(* IEC 61131-3 sources: daoli-st-library/DL_Base (part 7) *)

(* ---- FC_DL_RorEx.st ---- *)
(*==============================================================================
 * 组件名称 (Component)  : FC_DL_RorEx
 * 所属子库 (Sublibrary) : DL_Base
 * 当前版本 (Version)    : 1.0.0
 * 兼容性   (Platform)   : CODESYS 3.5 / TwinCAT 3 / 汇川 InoProShop / Machine Expert
 *                         仅依赖 Standard.library 的 SHL / SHR 内建函数，
 *                         循环语义由移位合成显式构造，无厂商 ROR 方言依赖
 * 功能一句话 (Summary)  : 循环右移防御包装：移位量对位宽取模归一后再循环，
 *                         杜绝平台相关行为，循环位不丢。
 * 功能描述 (Function)   : 对被移位位串按移位量 nN 循环右移。归一策略写死：
 *                         nN 先 MOD 32 归一到 0 到 31（nN 为 USINT 天然非负，
 *                         禁用 MOD 对负数的平台歧义取余的前提由类型系统保证）；
 *                         归一后 nN = 0 直接返回原值（整圈等价于不动，不置码）；
 *                         归一后 1 到 31 用「右移 nN OR 左移 (32 − nN)」位合成
 *                         构造循环语义，两个合成移位量均严格落在 1 到 31 安全域。
 * 溯源     (Origin)     : IEC 61131-3 标准语义的道莅防御性实现
 *                         （接口语义由 IEC 61131-3 定义，clean-room 重写，
 *                         参考公开标准条款）
 * 支持位宽 (Width Note) : 本件按 DWORD（32 位）主类型实现，仅支持 32 位位串；
 *                         BYTE / WORD 调用方先显式转换到 DWORD 后调用，再按需
 *                         截回原位宽（头注释显式声明，不做 ANY_BIT 泛型）。
 * 类型裁定 (Type Note)  : 码位段 16#0001_xxxx 为全库共享 32 位段，WORD 容量不足，
 *                         故 uDiag 采用 UDINT 承载（与库内 uErrorId : UDINT 惯例一致）
 * 依赖     (Depends)    : 无 DL_ 内部依赖；Standard.library: SHL / SHR
 * 红线自检 (Redline)    : R1 ✓ 零全局变量与外部变量引用 ｜ R2 ✓ 零物理 IO 地址直写
 *                         R3 ✓ 纯 IEC 61131-3 ｜ R4 ✓ 移位量 MOD 归一（合成移位
 *                         量恒在 1 到 31 安全域）｜ R5 ✓ 全变量中英双语同行注释
 *                         R6 N/A（纯函数，无 CASE/ENUM 状态机，按批 1 口径标 N/A）
 *                         R7 N/A（FC 为纯函数，无实例调用，头注释显式说明）
 * 防御行为声明 (Defense): ① 归一先行：nN ≥ 32 时先 MOD 32 归一并置信息码
 *                           16#0001_0159（已归一提示），归一后绝不出现 ≥ 位宽
 *                           的移位量，杜绝平台对超宽循环移位的歧义行为；
 *                         ② nN 为 USINT 类型天然非负，MOD 只作用于非负域，
 *                           负数取余的平台歧义（如商向零取整方向不一）从类型
 *                           系统层面被排除，该前提已在头注释写死；
 *                         ③ 归一后 nN = 0 直接返回原值且不置码（整圈无事件）；
 *                         ④ 位合成用「SHR(uIn, nN) OR SHL(uIn, 32 − nN)」，
 *                           nN 归一后为 1 到 31，故 32 − nN 恒为 1 到 31，
 *                           两个移位量均不触碰「移位量 = 位宽」禁区，循环位不丢；
 *                         ⑤ 32（位宽）提为只读常量，禁魔法数。
 * 修订历史 (Revision)   :
 *   2026-11-16  v1.0.0  首版入库（R14 批 3 · T0 快车道）
 *============================================================================*)
FUNCTION FC_DL_RorEx : DWORD
VAR_INPUT
    uIn : DWORD;   // 被循环移位位串 [位] / Bit string to be rotated
    nN  : USINT;   // 移位量 [bit]，USINT 天然非负，MOD 仅作用于非负域 / Shift amount [bit], USINT is non-negative, MOD applied on the non-negative domain only
END_VAR
VAR_OUTPUT
    uDiag : UDINT; // 诊断字，16#0001_0159=移位量已 MOD 32 归一，0=无事件 / Diag word, 16#0001_0159=shift amount reduced by MOD 32, 0=no event
END_VAR
VAR
    nNorm : USINT; // 归一后移位量 [bit]，域 0 到 31 / Normalized shift amount [bit], range 0 to 31
END_VAR
VAR CONSTANT
    DL_RR_WIDTH : USINT := 32;  // 位宽常量 [bit]，MOD 归一与合成移位共用 / Width constant [bit], shared by MOD normalization and composite shifts
END_VAR

(*------------------------------------------------------------------------------
 * 段 1｜输出与诊断预置：先归零，任何路径都不会留下脏诊断
 *      Pre-set the output and diag so no path ever leaves a stale diag
 *-----------------------------------------------------------------------------*)
FC_DL_RorEx := 16#0000_0000;   // 返回值预置全零 [位串] / Preset return value to all zero
uDiag       := 16#0000_0000;   // 诊断字预置无事件 / Preset diag word to no event
nNorm       := 0;              // 归一移位量预置 [bit] / Preset normalized shift to zero [bit]

(*------------------------------------------------------------------------------
 * 段 2｜移位量归一（防御声明①②）：nN MOD 32 归一到 0 到 31；
 *      nN 为 USINT 非负域，MOD 结果即数学取模，无负数取余歧义；
 *      nN ≥ 32 置信息码提示已归一（归一是正常防御行为，非故障）
 *      Shift-amount normalization (defense notes 1 and 2): nN MOD 32 reduces
 *      to 0 to 31; a reduction raises the informational code, not a fault
 *-----------------------------------------------------------------------------*)
IF nN >= DL_RR_WIDTH THEN
    nNorm := nN MOD DL_RR_WIDTH;   // 超宽归一：MOD 32 取模 [bit] / Oversized normalization: MOD 32 [bit]
    uDiag := 16#0001_0159;         // 信息码：移位量已 MOD 32 归一 / Informational: shift amount reduced by MOD 32
ELSE
    nNorm := nN;                   // 域内直通 [bit] / In-domain pass-through [bit]
END_IF

(*------------------------------------------------------------------------------
 * 段 3｜循环移位主体（防御声明③④）：归一后 0 整圈直通原值；
 *      1 到 31 用右移与左移位合成，合成移位量恒在安全域，循环位不丢
 *      Rotation body (defense notes 3 and 4): normalized zero returns as is;
 *      one to thirty one composes SHR and SHL, both amounts stay in the safe
 *      domain so no bit is ever lost
 *-----------------------------------------------------------------------------*)
IF nNorm = 0 THEN
    FC_DL_RorEx := uIn;   // 整圈（或 0 位）等价于原值直通 [位串] / A full turn (or zero shift) returns the input unchanged
ELSE
    FC_DL_RorEx := SHR(uIn, nNorm) OR SHL(uIn, DL_RR_WIDTH - nNorm);   // 位合成循环右移 [位串] / Composite rotate right
END_IF
END_FUNCTION

(* ---- FC_DL_RorLwordEx.st ---- *)
(*
    FC_DL_RorLwordEx —— LWORD 循环右移（MOD 64 归一）
    ------------------------------------------------------------------
    分类      : DL_Base / BitString
    前缀      : FC_DL_
    版本      : 1.0.0
    溯源      : IEC 61131-3 标准语义的道莅防御性实现
                （接口语义由 IEC 61131-3 定义，内部委托平台内建 ROR，
                  外围统一错误码 / 钳位 / 双语文档；clean-room 重写，
                  未复制任何闭源厂商源码，参考实现仅限 MIT/Apache 许可）
    平台      : 纯 IEC 61131-3，CODESYS / TwinCAT / InoProShop 通用
    作者      : 道莅代码库 · PLC编程专家（R17）
    ------------------------------------------------------------------
    功能说明  : LWORD 位串循环右移防御包装：移位量 nN 大于等于 64（位宽）时按 MOD 64 归一，
                并置信息级 16#0001_020C（与循环左移件同口径，与左移/右移件的「超宽置零」刻意相反）；
                归一后移位量为 0 时直接输出原值，不调用内建 ROR；
                域内委托平台内建 ROR，不重实现移位内核；
                MOD 除子为常量 64（编译期恒非零），结构性满足除法前判除子非零红线；
                钳位方向：移位量按位宽取模归一（0~63），结果位宽严格保持 64 位。
    错误码    : 16#0001_020C 移位量 ≥ 64（位宽），已按 MOD 64 归一——信息级，正常防御
                16#0001_020D 预留禁用（信息级，不得挪用）
                16#0001_0300 预留禁用（故障级，不得挪用）
                16#0001_0301 预留禁用（故障级，不得挪用）
                16#0001_0302 预留禁用（故障级，不得挪用）
    状态机    : R6 标注 N/A —— 本组件为纯函数无顺序状态机，无 CASE 可写，非法状态不可能出现，故以本节说明替代 ELSE 兜底
    修订记录  : 2026-11-16 v1.0.0 首次入库（R17）
*)
FUNCTION FC_DL_RorLwordEx : LWORD
VAR_INPUT
    uIn : LWORD; // 被循环移位位串 [位] / bit string to be rotated [bit]
    nN  : USINT; // 循环移位量 [bit]，USINT 天然非负，范围 0~255 / rotate amount [bit], USINT is non-negative by type, range 0..255
END_VAR
VAR_OUTPUT
    eErr   : UDINT; // 错误码，0=正常 / error id, 0=ok
    bError : BOOL;  // 是否出错，eErr 非 0 时为 TRUE / error flag, TRUE when eErr is nonzero
    bValid : BOOL;  // 输出是否有效可用 / output valid flag
END_VAR
VAR CONSTANT
    DL_LW_WIDTH : USINT := 64; // LWORD 位宽常量，兼作 MOD 除子（编译期恒非零） [bit] / LWORD width constant, also the MOD divisor, never zero [bit]
END_VAR
VAR
    nShift : USINT; // 归一后的实际移位量 0~63 [bit] / normalized shift amount 0..63 [bit]
END_VAR

// 段 1｜输出与错误状态预置 / segment 1, preset output and error status
FC_DL_RorLwordEx := uIn; // 输出预置为原值（零移位等价语义），任何路径不留脏值 [位串] / preset output to the input, the zero-shift identity, no stale value on any path [bit string]
eErr   := 0;     // 预置无错误 / preset no error
bError := FALSE; // 预置无故障（本件无故障级路径） / preset no fault, no fault-level path here
bValid := FALSE; // 预置输出无效，通过归一后置位 / preset invalid, set TRUE after normalization

// 段 2｜移位量归一（MOD 位宽） / segment 2, shift amount normalization (modulo width)
nShift := nN; // 默认按原移位量直通 [bit] / pass the original shift amount through by default [bit]
IF nN >= DL_LW_WIDTH THEN // 循环移位对位宽取模仍等价，故归一而非置零 [bit] / rotate modulo the width stays equivalent, so normalize instead of zeroing [bit]
    nShift := nN MOD DL_LW_WIDTH; // 除子为编译期常量 64，恒非零 [bit] / divisor is the compile-time constant 64, never zero [bit]
    eErr := 16#0001_020C;         // 信息级：移位量已归一，正常防御 / info level: shift amount normalized, normal defence
ELSE
    eErr := 0;                    // 未超宽，无记录 / not oversized, nothing recorded
END_IF

// 段 3｜零移位量与域内委托循环移位（末段） / segment 3, zero-shift pass-through and in-domain delegated rotate (final)
IF nShift = 0 THEN
    FC_DL_RorLwordEx := uIn; // 零移位量直接输出原值，规避内建 ROR 的平台差异 [位串] / zero shift passes the input through, avoiding platform differences of built-in ROR [bit string]
ELSE
    FC_DL_RorLwordEx := ROR(uIn, nShift); // 域内委托平台内建 ROR，不重实现移位内核 [位串] / in-domain delegate to built-in ROR, shift kernel not re-implemented [bit string]
END_IF
bError := FALSE; // 信息级不置故障 / info level never raises fault
bValid := TRUE;  // 归一后输出有效可用 / output is valid after normalization
END_FUNCTION

(* ---- FC_DL_SaturateDiv.st ---- *)
(*
  ==================================================================
  组件名 Component  : FC_DL_SaturateDiv
  分类   Category   : DL_Base
  前缀   Naming     : FC_DL_ ｜ b/n/u/f/t/e/st 类型前缀制（R265）
  码位   Code ID    : 16#0001_0647（信息级）｜ 16#0001_0648 / 0649 / 064A（故障级）
  版本   Version    : 1.0.0
  复杂度 Complexity  : 中
  功能   Purpose    : LINT 宽域饱和除法：nOut = clamp(nNum ÷ nDen, nLo, nHi)，判据有序
                      （除零 → MIN÷-1 → 正常除 → 域钳），整数商向零截断。
  开源溯源 Origin    : IEC 61131-3 标准语义的道莅防御性实现（clean-room，无第三方代码行）
  许可证 License    : MIT
  参考   Reference  : IEC 61131-3:2013 §6.6.2 算术运算符（整数除法，商向零截断）
  平台   Platform   : 纯 IEC 61131-3（仅四则与比较），CODESYS / TwinCAT 3 / InoProShop 通用
  依赖   Depends    : 仅 Standard.library（无库调用）
  分工声明 Split     : FC_DL_DivDintSafeChk 为「安全除 + 商出口 + 布尔返回」的判据件
                      （DINT 域、无钳位域）；FC_DL_DivLrealSafe 为浮点域安全除；
                      本件为宽域（LINT）饱和除，带钳位域与三段标志。三者边界：
                      需要「除零仅判不钳」用前者，需要「浮点除法」用中者，
                      需要「整数宽域 + 钳位域 + 溢出标志」用本件（R216 双向互引）。
  归属 Ownership     : 本件无 TYPE 声明，全部引脚为 IEC 标准原生类型。
  ------------------------------------------------------------------
  边界 Boundary     :
                      一 判据严格有序：① 除数为零 → 早退（禁走钳位，钳位会把非法
                         结果伪装成合法边界）；② MIN ÷ -1 → 溢出钳 nHi；③ 正常除；
                         ④ 结果钳域 [nLo, nHi]；
                      二 商向零截断（IEC 语义）：-7 ÷ 2 = -3 而非 -4；本件不做四舍五入，
                         工程舍入口径归 FC_DL_RoundSat，有效位舍入归 FC_DL_RoundSigFigs；
                      三 nLo > nHi 判组态故障并返回 FALSE（与 FC_DL_SaturateMul、
                         FC_DL_RealToIntSat 同口径，三件一致，禁静默交换）；
                      四 纯函数：无记忆量、无定时器、无边沿实例，每调用重算。
  错误码 Codes      :
    16#0001_0647【信息级】结果被域 [nLo, nHi] 钳位（未溢出、未除零，bValid = TRUE）
    16#0001_0648【故障级】除数为零（nOut = 0，bValid = FALSE，早退不走钳位）
    16#0001_0649【故障级】MIN ÷ -1 溢出（nOut 钳 nHi，bOvF = TRUE）
    16#0001_064A【故障级】组态非法 nLo > nHi（判故障返回 FALSE，nOut = 0）
  码位反证 Note     :
    0648 不可并入 0647：除零结果与钳位结果在数值出口上同为边界值或零，上游无法由
    nOut 与 bClamped 组合区分「输入非法」与「输入合法但被限幅」，两码必需（R90）。
  验收 Acceptance   :
    算法已证（脚本）：未跑 ｜ 编译器已证（三平台）：未跑
    V1 5 ÷ 0 → 0、bDivZero = TRUE、bValid = FALSE、码 0648（不走钳位）
    V2 MIN ÷ -1 → nHi、bOvF = TRUE、码 0649
    V3 MIN ÷ 1 → MIN 精确
    V4 1 ÷ MIN → 0，bClamped = FALSE（未触钳位，仅截断）
    V5 -7 ÷ 2 → -3（向零截断，非 -4）
    V6 nLo > nHi → 码 064A、返回 FALSE
    V7 100 ÷ 3 = 33（截断）、域 [0, 20] → bClamped = TRUE、码 0647、bValid = TRUE
    V8 MIN ÷ -3 → 正常除（除子非 -1）不溢出
  修订记录 Revision  :
    2026-11-21  v1.0.0  R62 首版（批 1 · 序号 2）
  ==================================================================
*)
FUNCTION FC_DL_SaturateDiv : BOOL
VAR_INPUT
    nNum : LINT; // 被除数 [−]，完整 LINT 域 / the dividend over the full LINT domain
    nDen : LINT; // 除数 [−]，零为非法（判故障）/ the divisor, zero is illegal and raises a fault
    nLo  : LINT; // 输出钳位域下界 [−] / the output clamp lower bound
    nHi  : LINT; // 输出钳位域上界 [−] / the output clamp upper bound
END_VAR
VAR_OUTPUT
    nOut     : LINT;  // 钳位后商 [−] / the clamped quotient
    bDivZero : BOOL;  // 除数为零 [-] / the divisor is zero
    bOvF     : BOOL;  // 溢出发生（MIN ÷ -1）[-] / an overflow happened on MIN divided by minus one
    bClamped : BOOL;  // 钳位生效（含纯域钳）[-] / the clamp took effect, domain clamp included
    bValid   : BOOL;  // 输出可用（除零与组态故障为 FALSE）[-] / the output is usable
    eErr     : UDINT; // 错误码，0 = 正常 / the error code, zero is ok
    bError   : BOOL;  // 故障标志，故障级码同拍置位（R45 配对）/ the fault flag, raised with a fault level code
END_VAR
VAR
    liQuot : LINT := 0; // 域内商中间量 [−] / the in-domain quotient intermediate
END_VAR  // R64 结构补齐：VAR 段缺失的 END_VAR（门禁机械修复）
VAR CONSTANT
    DL_SDIV_MAX : LINT := 9223372036854775807;      // LINT 可表达上界 [−]，独立命名不与乘法件冲突 / the expressible LINT ceiling under its own name
    DL_SDIV_MIN : LINT := -9223372036854775807 - 1; // LINT 可表达下界 [−]，以上界相反数减一表达 / the expressible LINT floor written as the negated ceiling minus one
    DL_SDIV_ZERO : LINT := 0;                       // 有符号零常量 [−] / the signed zero constant
    DL_SDIV_NEG1 : LINT := -1;                      // 负一常量 [−]，MIN ÷ -1 判据用 / the minus one constant for the MIN divided by minus one criterion
END_VAR

// 段 1｜返回值与全部出口预置安全值（R45 四段式第一段）/ segment 1, preset every outlet to its safe value
FC_DL_SaturateDiv := FALSE; // 返回值预置假 / preset the return false
nOut := DL_SDIV_ZERO; // 结果预置零 [−] / preset the quotient zero
bDivZero := FALSE; // 除零标志预置假 / preset the divide by zero flag false
bOvF := FALSE; // 溢出标志预置假 / preset the overflow flag false
bClamped := FALSE; // 钳位标志预置假 / preset the clamp flag false
bValid := FALSE; // 可用标志预置假，过闸后置位 / preset the validity false, raised after the gates
eErr := 16#0000_0000; // 错误码预置正常 / preset the code to ok
bError := FALSE; // 故障标志预置假 / preset the fault flag false
liQuot := DL_SDIV_ZERO; // 商中间量清零 [−] / clear the quotient intermediate

// 段 2｜组态域闸：nLo > nHi 判故障早退（边界三，三件同口径）/ segment 2, the configuration gate, a reversed domain is a fault
IF nLo > nHi THEN // 钳位域反序 / the clamp domain is reversed
    eErr := 16#0001_064A; // 故障级：组态非法 nLo > nHi / fault grade, the reversed clamp domain
    bError := TRUE; // 同拍置故障标志（R45 配对）/ raise the fault flag on the same scan
    bValid := FALSE; // 输出不可用 / the output is not usable
    nOut := DL_SDIV_ZERO; // 确定缺省值零 [−] / the deterministic default of zero
    RETURN; // 早退 / early return
END_IF

// 段 3｜判据①除数为零：早退，绝不行钳位（边界一，钳位会把非法伪装成合法边界）/ segment 3, the divisor zero gate, clamped never runs
IF nDen = DL_SDIV_ZERO THEN // 除数为零 / the divisor is zero
    bDivZero := TRUE; // 置除零标志 / raise the divide by zero flag
    nOut := DL_SDIV_ZERO; // 确定缺省值零 [−] / the deterministic default of zero
    eErr := 16#0001_0648; // 故障级：除数为零 / fault grade, the divisor is zero
    bError := TRUE; // 同拍置故障标志（R45 配对）/ raise the fault flag on the same scan
    bValid := FALSE; // 输出不可用 / the output is not usable
    RETURN; // 早退，不做任何除法与钳位 / early return without any division or clamping
END_IF

// 段 4｜判据②MIN ÷ -1 溢出（MIN 的绝对值不可表示，先除必回绕）/ segment 4, the MIN divided by minus one overflow
IF (nNum = DL_SDIV_MIN) AND (nDen = DL_SDIV_NEG1) THEN // 极限组合 / the limit combination
    bOvF := TRUE; // 置溢出标志（禁回绕成 MIN）/ raise the overflow flag instead of wrapping to MIN
    bClamped := TRUE; // 钳位已生效 / the clamp took effect
    nOut := nHi; // 正溢出按符号钳上界 [−] / a positive overflow clamps to the upper bound by sign
    eErr := 16#0001_0649; // 故障级：MIN ÷ -1 溢出 / fault grade, the MIN divided by minus one overflow
    bError := TRUE; // 同拍置故障标志（R45 配对）/ raise the fault flag on the same scan
    bValid := FALSE; // 输出不可用 / the output is not usable
    RETURN; // 早退 / early return
END_IF

// 段 5｜判据③正常除：整数商向零截断（边界二，IEC 语义，-7 ÷ 2 = -3）/ segment 5, the normal division with the quotient truncated toward zero
IF nNum = DL_SDIV_ZERO THEN // 零被除数：商确为零，免一次除法 / a zero dividend gives an exact zero quotient, no division needed
    liQuot := DL_SDIV_ZERO; // 商为零 [−] / the quotient is zero
ELSE // 非零被除数才真除（除子已在段 3 证非零）/ the real division only for a nonzero dividend, the divisor is proven nonzero
    liQuot := nNum / nDen; // 向零截断（-7 ÷ 2 = -3，非 -4）[−] / truncated toward zero, minus seven over two gives minus three
END_IF

// 段 6｜判据④统一域钳（零被除数与正常除共用同一出口，R94）/ segment 6, the unified domain clamp shared by both paths
IF liQuot > nHi THEN // 超上界 / above the ceiling
    nOut := nHi; // 钳上界 [−] / clamp to the ceiling
    bClamped := TRUE; // 置钳位标志 / raise the clamp flag
ELSIF liQuot < nLo THEN // 超下界 / below the floor
    nOut := nLo; // 钳下界 [−] / clamp to the floor
    bClamped := TRUE; // 置钳位标志 / raise the clamp flag
ELSE // 域内 / inside the domain
    nOut := liQuot; // 直出商 [−] / pass the quotient through
END_IF

// 段 7｜信息级钳位码与可用位（纯域钳不置 bError，R285）/ segment 7, the informational clamp code without a fault flag
IF bClamped THEN // 发生纯域钳 / a pure domain clamp happened
    eErr := 16#0001_0647; // 信息级：结果被域钳位 / informational, the result was clamped to the domain
END_IF
bValid := TRUE; // 域内或钳位输出均可用 / an in-domain or clamped output is usable
FC_DL_SaturateDiv := TRUE; // 返回成功 / return success
END_FUNCTION

(* ---- FC_DL_SaturateMul.st ---- *)
(*
  ==================================================================
  组件名 Component  : FC_DL_SaturateMul
  分类   Category   : DL_Base
  前缀   Naming     : FC_DL_ ｜ b/n/u/f/t/e/st 类型前缀制（R265）
  码位   Code ID    : 16#0001_0644（信息级）｜ 16#0001_0645（故障级）｜ 16#0001_0646（故障级）
  版本   Version    : 1.0.0
  复杂度 Complexity  : 中
  功能   Purpose    : LINT 宽域饱和乘法：nOut = clamp(nA × nB, nLo, nHi)，溢出前判定，
                      bOvF（溢出）与 bClamped（钳位已生效）两标志语义可分。
  开源溯源 Origin    : IEC 61131-3 标准语义的道莅防御性实现（clean-room，无第三方代码行）
  许可证 License    : MIT
  参考   Reference  : IEC 61131-3:2013 §6.6.2 算术运算符（整数乘法）与 §6.6.5 类型转换语义
  平台   Platform   : 纯 IEC 61131-3（仅四则与比较），CODESYS / TwinCAT 3 / InoProShop 通用
  依赖   Depends    : 仅 Standard.library（无库调用）
  分工声明 Split     : 与 FC_DL_SaturateAdd（加）/ FC_DL_SaturateSub（减）构成「加/减/乘」
                      三件族，除法则由 FC_DL_SaturateDiv 承载；FC_DL_SaturateAdd 未覆盖
                      乘法（其模式枚举只有加与减），故本件不可省（R216 双向互引）。
  归属 Ownership     : 本件无 TYPE 声明，全部引脚为 IEC 标准原生类型。
  ------------------------------------------------------------------
  边界 Boundary     :
                      一 溢出前判定（禁先乘后判）：按四个象限分别与「域上界 ÷ 另一因子」
                         比较，比较式内只出现除法，不出现裸乘法，浮点无关、全整数精确；
                      二 MIN × -1 单独直判：MIN 的绝对值不可表示，先乘必回绕成 MIN 而
                         令「结果 < 0」误判为负溢出，故本组合在乘法之前直接判正溢出；
                      三 零因子优先：nA = 0 或 nB = 0 时积恒为 0，不做任何除法预判
                         （同时消灭预判式里的除零路径）；
                      四 nLo > nHi 判组态故障并返回 FALSE（与 FC_DL_SaturateDiv、
                         FC_DL_RealToIntSat 同口径，三件一致，禁静默交换）；
                      五 溢出与域钳两标志可分：溢出 → bOvF = TRUE 且 nOut 直达 nHi/nLo；
                         未溢出仅域钳 → bClamped = TRUE 且 bOvF = FALSE；
                      六 纯函数：无记忆量、无定时器、无边沿实例，每调用重算。
  错误码 Codes      :
    16#0001_0644【信息级】结果被域 [nLo, nHi] 钳位（未溢出，bClamped = TRUE，bValid = TRUE）
    16#0001_0645【故障级】乘法溢出（bOvF = TRUE，nOut 已按积符号钳到 nHi 或 nLo）
    16#0001_0646【故障级】组态非法 nLo > nHi（判故障返回 FALSE，nOut = 0）
  码位反证 Note     :
    0644 与 0645 不可合并：溢出与域钳在「结果数值」上不可观测区分（两者都输出边界值），
    仅靠返回值加 bValid 也无法分解（两者 bValid 不同，但 bOvF 语义才是上游限幅判据），
    故两码必需（R90 反证句：现有输出组合无法唯一还原该场景）。
  验收 Acceptance   :
    算法已证（脚本）：未跑 ｜ 编译器已证（三平台）：未跑
    V1 MAX × 2 → nOut = nHi、bOvF = TRUE、码 0645
    V2 MIN × -1 → nOut = nHi、bOvF = TRUE（禁回绕成 MIN）
    V3 MIN × 0 → 0 且 bOvF = FALSE
    V4 MIN × 1 → MIN 精确（无溢出、无钳位）
    V5 -3 × 5 → -15 精确
    V6 nLo > nHi → 码 0646、bError = TRUE、返回 FALSE
    V7 nLo = nHi = 100、积 = 200 → bClamped = TRUE 且 bOvF = FALSE（两标志可分）
    V8 nA = 0、nB = MIN → 0（零因子早于预判，无除零）
  修订记录 Revision  :
    2026-11-21  v1.0.0  R62 首版（批 1 · 序号 1）
  ==================================================================
*)
FUNCTION FC_DL_SaturateMul : BOOL
VAR_INPUT
    nA   : LINT; // 被乘数 [−]，完整 LINT 域 / the multiplicand over the full LINT domain
    nB   : LINT; // 乘数 [−]，完整 LINT 域 / the multiplier over the full LINT domain
    nLo  : LINT; // 输出钳位域下界 [−] / the output clamp lower bound
    nHi  : LINT; // 输出钳位域上界 [−] / the output clamp upper bound
END_VAR
VAR_OUTPUT
    nOut     : LINT;  // 钳位后结果 [−] / the clamped product
    bOvF     : BOOL;  // 乘法溢出发生（钳位已生效）[-] / a multiplicative overflow happened
    bClamped : BOOL;  // 钳位生效（含纯域钳，未溢出）[-] / the clamp took effect, domain clamp included
    bValid   : BOOL;  // 输出可用（溢出与组态故障为 FALSE）[-] / the output is usable
    eErr     : UDINT; // 错误码，0 = 正常 / the error code, zero is ok
    bError   : BOOL;  // 故障标志，故障级码同拍置位（R45 配对）/ the fault flag, raised with a fault level code
END_VAR
VAR
    liProd : LINT := 0; // 域内乘积中间量 [−] / the in-domain product intermediate
END_VAR  // R64 结构补齐：VAR 段缺失的 END_VAR（门禁机械修复）
VAR CONSTANT
    DL_SMUL_MAX : LINT := 9223372036854775807;      // LINT 可表达上界 [−]，即 2^63−1 / the expressible LINT ceiling, two to the sixty third minus one
    DL_SMUL_MIN : LINT := -9223372036854775807 - 1; // LINT 可表达下界 [−]，以上界相反数减一表达，防字面量解析溢出 / the expressible LINT floor, written as the negated ceiling minus one to avoid a literal parse overflow
    DL_SMUL_ZERO : LINT := 0;                       // 有符号零常量 [−]，避免裸字面量 / the signed zero constant
    DL_SMUL_NEG1 : LINT := -1;                      // 负一常量 [−]，MIN × -1 判据用 / the minus one constant for the MIN times minus one criterion
END_VAR

// 段 1｜返回值与全部出口预置安全值（R45 四段式第一段）/ segment 1, preset every outlet to its safe value
FC_DL_SaturateMul := FALSE; // 返回值预置假 / preset the return false
nOut := DL_SMUL_ZERO; // 结果预置零 [−] / preset the product zero
bOvF := FALSE; // 溢出标志预置假 / preset the overflow flag false
bClamped := FALSE; // 钳位标志预置假 / preset the clamp flag false
bValid := FALSE; // 可用标志预置假，过闸后置位 / preset the validity false, raised after the gates
eErr := 16#0000_0000; // 错误码预置正常 / preset the code to ok
bError := FALSE; // 故障标志预置假 / preset the fault flag false
liProd := DL_SMUL_ZERO; // 乘积中间量清零 [−] / clear the product intermediate

// 段 2｜组态域闸：nLo > nHi 判故障早退（边界四，三件同口径）/ segment 2, the configuration gate, a reversed domain is a fault
IF nLo > nHi THEN // 钳位域反序 / the clamp domain is reversed
    eErr := 16#0001_0646; // 故障级：组态非法 nLo > nHi / fault grade, the reversed clamp domain
    bError := TRUE; // 同拍置故障标志（R45 配对）/ raise the fault flag on the same scan
    bValid := FALSE; // 输出不可用 / the output is not usable
    nOut := DL_SMUL_ZERO; // 确定缺省值零 [−] / the deterministic default of zero
    RETURN; // 早退，不再触碰乘法 / early return, the multiplication is never touched
END_IF

// 段 3｜零因子优先：积恒为零，且消灭后续预判式的除零路径（边界三）/ segment 3, the zero factor comes first and removes every division by zero
IF (nA = DL_SMUL_ZERO) OR (nB = DL_SMUL_ZERO) THEN // 任一因子为零 / either factor is zero
    liProd := DL_SMUL_ZERO; // 积确定为零 [−] / the product is exactly zero
ELSE // 双因子非零才做溢出预判 / the overflow pre-check runs only with two nonzero factors
    // 段 4｜MIN × -1 直判正溢出（边界二）：MIN 绝对值不可表示，先乘会回绕成 MIN / segment 4, the direct check of MIN times minus one
    IF ((nA = DL_SMUL_MIN) AND (nB = DL_SMUL_NEG1)) OR ((nB = DL_SMUL_MIN) AND (nA = DL_SMUL_NEG1)) THEN // 极限组合 / the limit combination
        bOvF := TRUE; // 置溢出标志（禁回绕成 MIN）/ raise the overflow flag instead of wrapping to MIN
        bClamped := TRUE; // 钳位已生效 / the clamp took effect
        nOut := nHi; // 正溢出按符号钳上界 [−] / a positive overflow clamps to the upper bound by sign
        eErr := 16#0001_0645; // 故障级：乘法溢出 / fault grade, a multiplicative overflow
        bError := TRUE; // 同拍置故障标志（R45 配对）/ raise the fault flag on the same scan
        bValid := FALSE; // 输出不可用（结果是伪造边界）/ the output is not usable, the boundary is fabricated
        RETURN; // 早退 / early return
    END_IF
    // 段 5｜四象限溢出预判（边界一）：比较式内只有除法，没有裸乘法 / segment 5, the four quadrant pre-check with divisions only
    IF (nA > DL_SMUL_ZERO) AND (nB > DL_SMUL_ZERO) THEN // 正正象限 / the positive positive quadrant
        IF nA > (DL_SMUL_MAX / nB) THEN // 超上界预判（nB ≥ 1，除子安全）/ the ceiling pre-check with a safe divisor
            bOvF := TRUE; // 置溢出标志 / raise the overflow flag
            bClamped := TRUE; // 钳位已生效 / the clamp took effect
            nOut := nHi; // 正溢出钳上界 [−] / a positive overflow clamps to the upper bound
        END_IF
    ELSIF (nA < DL_SMUL_ZERO) AND (nB < DL_SMUL_ZERO) THEN // 负负象限（积为正）/ the negative negative quadrant, a positive product
        IF nA < (DL_SMUL_MAX / nB) THEN // 超上界预判（MAX ÷ 负数为负，直比不失号）/ the ceiling pre-check against a negative quotient
            bOvF := TRUE; // 置溢出标志 / raise the overflow flag
            bClamped := TRUE; // 钳位已生效 / the clamp took effect
            nOut := nHi; // 正溢出钳上界 [−] / a positive overflow clamps to the upper bound
        END_IF
    ELSIF (nA > DL_SMUL_ZERO) AND (nB < DL_SMUL_ZERO) THEN // 正负象限（积为负）/ the positive negative quadrant, a negative product
        IF nB < (DL_SMUL_MIN / nA) THEN // 超下界预判（nA ≥ 1，除子安全）/ the floor pre-check with a safe divisor
            bOvF := TRUE; // 置溢出标志 / raise the overflow flag
            bClamped := TRUE; // 钳位已生效 / the clamp took effect
            nOut := nLo; // 负溢出钳下界 [−] / a negative overflow clamps to the lower bound
        END_IF
    ELSE // 负正象限（积为负）/ the negative positive quadrant, a negative product
        IF nA < (DL_SMUL_MIN / nB) THEN // 超下界预判（nB ≥ 1，除子安全）/ the floor pre-check with a safe divisor
            bOvF := TRUE; // 置溢出标志 / raise the overflow flag
            bClamped := TRUE; // 钳位已生效 / the clamp took effect
            nOut := nLo; // 负溢出钳下界 [−] / a negative overflow clamps to the lower bound
        END_IF
    END_IF
    IF bOvF THEN // 已判溢出：结果已直达边界，跳过域钳 / an overflow already reached the boundary, the domain clamp is skipped
        eErr := 16#0001_0645; // 故障级：乘法溢出 / fault grade, a multiplicative overflow
        bError := TRUE; // 同拍置故障标志（R45 配对）/ raise the fault flag on the same scan
        bValid := FALSE; // 输出不可用 / the output is not usable
        RETURN; // 早退 / early return
    END_IF
    liProd := nA * nB; // 预判通过后域内相乘（此时必不溢出）/ multiply after the pre-check passed, so no overflow can occur
END_IF

// 段 6｜统一域钳（零因子与域内积共用同一出口，R94 早退分支后处理一致）/ segment 6, the unified domain clamp shared by both paths
IF liProd > nHi THEN // 超上界 / above the ceiling
    nOut := nHi; // 钳上界 [−] / clamp to the ceiling
    bClamped := TRUE; // 置钳位标志 / raise the clamp flag
ELSIF liProd < nLo THEN // 超下界 / below the floor
    nOut := nLo; // 钳下界 [−] / clamp to the floor
    bClamped := TRUE; // 置钳位标志 / raise the clamp flag
ELSE // 域内 / inside the domain
    nOut := liProd; // 直出乘积 [−] / pass the product through
END_IF

// 段 7｜信息级钳位码与可用位（纯域钳不置 bError，R285 分级纪律）/ segment 7, the informational clamp code without a fault flag
IF bClamped THEN // 发生纯域钳（溢出已在段 5 早退）/ a pure domain clamp happened, overflow already returned earlier
    eErr := 16#0001_0644; // 信息级：结果被域钳位 / informational, the result was clamped to the domain
END_IF
bValid := TRUE; // 域内或钳位输出均可用 / an in-domain or clamped output is usable
FC_DL_SaturateMul := TRUE; // 返回成功 / return success
END_FUNCTION

(* ---- FC_DL_SaturateSub.st ---- *)
(*==============================================================================
 * 组件名称 (Component)  : FC_DL_SaturateSub
 * 所属子库 (Sublibrary) : DL_Base
 * 当前版本 (Version)    : 1.0.1
 * 兼容性   (Platform)   : CODESYS 3.5+ / TwinCAT 3 / 汇川 InoProShop / 施耐德 Machine Expert
 *                         仅依赖 Standard.library，零厂商私有库
 * 功能描述 (Function)   : 有符号整数（DINT）饱和减法原语：nResult = nMinuend - nSubtrahend，
 *                         结果若超出 DINT 可表域则钳位返回 DINT 域下限/上限，并经引用参数
 *                         bOverflow 置溢出标志；正常域 bOverflow := FALSE。
 *                         与 `FC_DL_SaturateAdd` 成对（那件管累加方向防回绕，本件管扣减方向
 *                         防回绕），实现独立、只对齐注释风格与引脚组织，不复制其实现。
 * 接口     (Interface)  : 输入 nMinuend 被减数、nSubtrahend 减数；
 *                         引用输出 bOverflow 溢出标志（REFERENCE TO BOOL，当拍写回）；
 *                         返回值 = 饱和后的差（DINT）。
 * 边界     (Boundary)   : ① **属主边界（写死）：本件只做单次减法饱和运算，不记忆任何跨拍状态、
 *                         不接管计数器/累积器语义**；调用方自持累积变量并按需调用本件。
 *                         ② 溢出判定采用「先判后算」跨域预判，禁止先算后判（先算后判时中间值
 *                         已回绕、溢出不可观测）：减数 > 0 时下溢预判式为
 *                         nMinuend < (DINT 下限 + 减数)；减数 < 0 时上溢预判式为
 *                         nMinuend > (DINT 上限 + 减数)。两个预判式中的加法结果均在 DINT
 *                         域内可表（下限+正数 ≤ 上限方向、上限+负数 ≥ -1），不产生新的回绕。
 *                         ③ 减数 = 0 时恒为直通拷贝，无溢出可能，bOverflow 恒 FALSE。
 *                         ④ 边界向量覆盖：MIN_INT - (-1)、MAX_INT - 负数、MIN_INT - 正数、
 *                         零减零，详见头注释修订记录所附验收向量。
 *                         ⑤ 零全局耦合（无 GVL / 无 VAR_EXTERNAL / 无物理地址）。
 * 分工声明 (Scope)      : 与 `FC_DL_SaturateAdd` 分工：累加方向防回绕归那件、扣减方向防回绕
 *                         归本件（余料核销、步进回退计数等减法域）；二者不互相调用。
 * 来源标签 (Source Tag) : 自研线（成对补口，公开饱和运算定义 clean-room）
 * 码表     (Codes)      : 本件不占用任何全局数字码位。出口为 DINT 差值 + BOOL 溢出标志；
 *                         数字码位待主控收口阶段统一派号。
 * 红线自检 (Redline)    : R1 ✓ 零 GVL/VAR_EXTERNAL ｜ R2 ✓ 零 %I/%Q/%M ｜ R3 ✓ 纯 IEC 61131-3
 *                         R4 ✓ 先判后算跨域预判 + 类型可表性反算 ｜ R5 ✓ 声明逐行同行双语注释
 *                         R6 N/A（纯函数无状态机） ｜ R7 N/A（无实例调用）
 * 修订历史 (Revision)   : 2026-11-20  v1.0.1  R50 返修 R5：头注释验收向量溢出
 *                         断言更正（实现不动）——原「MIN-(-1)=MIN 溢出」为误
 *                         断言：MIN−(−1) = −2147483647 在 DINT 域内可表，无
 *                         溢出（预判式 nMinuend > MAX−1 对 MIN 不成立，实现
 *                         行为正确）；更正为「MIN-(-1)=MIN+1 正常」。另
 *                         「MIN-1=MIN 溢出」复核成立（MIN−1 下溢钳 MIN）。
 *                         2026-11-20  v1.0.0  R48 首版（批次 1 · 序号 1）
 *                         验收向量：MAX-(-1)=MAX 溢出；MIN-1=MIN 溢出；
 *                         MIN-(-1)=-2147483647 正常（v1.0.1 更正）；0-0=0 正常；
 *                         MIN-MIN=0 正常；MAX-MIN=MAX 溢出。
 *==============================================================================*)

FUNCTION FC_DL_SaturateSub : DINT
VAR_INPUT
    nMinuend    : DINT;                // 被减数 [-] / Minuend of the subtraction
    nSubtrahend : DINT;                // 减数 [-] / Subtrahend of the subtraction
    bOverflow   : REFERENCE TO BOOL;   // 溢出标志（引用传参，当拍写回；TRUE=已钳位） [-] / Overflow flag, by-reference, TRUE when clamped
END_VAR
VAR CONSTANT
    DL_SBS_MIN : DINT := DINT#16#80000000;   // DINT 域下限（类型可表性下界；位型常量，非事件码） [-] / DINT lower bound, bit-pattern constant, not an event code
    DL_SBS_MAX : DINT := 2147483647;         // DINT 域上限（类型可表性上界） [-] / DINT upper bound
END_VAR

(* —— 先判后算：跨域预判溢出，杜绝中间值回绕不可观测 —— *)
bOverflow := FALSE;                                                      // 正常域缺省无溢出 / Default: no overflow
IF nSubtrahend > 0 THEN                                                  // 减数为正：只可能下溢 / Positive subtrahend: underflow only
    IF nMinuend < (DL_SBS_MIN + nSubtrahend) THEN                        // 预判式在 DINT 域内可表 / Pre-check stays representable in DINT
        bOverflow := TRUE;                                               // 下溢成立：置溢出标志 / Underflow: raise overflow flag
        FC_DL_SaturateSub := DL_SBS_MIN;                                 // 钳位返回 DINT 下限 / Clamp to DINT lower bound
        RETURN;                                                          // 早退，不做真实减法 / Early exit, skip the raw subtraction
    END_IF
ELSIF nSubtrahend < 0 THEN                                               // 减数为负：只可能上溢 / Negative subtrahend: overflow only
    IF nMinuend > (DL_SBS_MAX + nSubtrahend) THEN                        // 预判式在 DINT 域内可表 / Pre-check stays representable in DINT
        bOverflow := TRUE;                                               // 上溢成立：置溢出标志 / Overflow: raise overflow flag
        FC_DL_SaturateSub := DL_SBS_MAX;                                 // 钳位返回 DINT 上限 / Clamp to DINT upper bound
        RETURN;                                                          // 早退，不做真实减法 / Early exit, skip the raw subtraction
    END_IF
END_IF

FC_DL_SaturateSub := nMinuend - nSubtrahend;                             // 已证可表的正常域减法 / Subtraction proven representable

END_FUNCTION

(* ---- FC_DL_SevenSegBcdDecode.st ---- *)
(* ============================================================
   DL_Base / FC_DL_SevenSegBcdDecode ｜ v1.0.0 ｜ 2026-11-25
   功能：BCD 位（0~9）→ 七段段码。段位 bit0=a bit1=b bit2=c bit3=d bit4=e
         bit5=f bit6=g bit7=dp；bCommonAnode=TRUE 整字节取反（共阳低有效）
   边界：输入 > 9 → 全灭（共阴 16#00 / 共阳 16#FF）且 bValid=FALSE；
         小数点叠加不属本件（签名无 dp 引脚），由 FC_DL_SevenSegMinusFlagCalc 负责；
         本文件 16# 常量均为段掩码，非事件码位（R83 不入账）
   依赖：仅 IEC 61131-3（NOT） ｜ 溯源：DLF-C-SEVENSEG（内部原创线）
   ============================================================ *)
FUNCTION FC_DL_SevenSegBcdDecode : BOOL
VAR_INPUT
    uBcd         : BYTE;  // BCD 位值，域 0~9 [-] / BCD digit, domain zero to nine
    bCommonAnode : BOOL;  // TRUE=共阳低有效 / FALSE=共阴高有效 [-] / TRUE for common anode
END_VAR
VAR_OUTPUT
    uSegCode : BYTE;  // 七段段码（含极性，不含 dp）[-] / Segment code with polarity, without dp
    bValid   : BOOL;  // 输入在 BCD 域内 [-] / Input inside the BCD domain
END_VAR
VAR
    _uRaw : BYTE;  // 共阴原始段码 [-] / Raw common cathode code
END_VAR

(* 段 0：出口预置安全侧（全灭按极性，N3） *)
FC_DL_SevenSegBcdDecode := FALSE;
_uRaw := 16#00;
bValid := FALSE;
IF bCommonAnode THEN uSegCode := 16#FF; ELSE uSegCode := 16#00; END_IF

(* 段 1：BCD 域闸（> 9 保持全灭，不做隐式回绕） *)
IF uBcd > 9 THEN RETURN; END_IF

(* 段 2：字形查表（段掩码常量，非码位） *)
CASE uBcd OF
0: _uRaw := 16#3F;   // 段 abcdef / Segments a to f
1: _uRaw := 16#06;   // 段 bc / Segments b and c
2: _uRaw := 16#5B;   // 段 abdeg / Segments a b d e g
3: _uRaw := 16#4F;   // 段 abcdg / Segments a b c d g
4: _uRaw := 16#66;   // 段 bcfg / Segments b c f g
5: _uRaw := 16#6D;   // 段 acdfg / Segments a c d f g
6: _uRaw := 16#7D;   // 段 acdefg / Segments a c d e f g
7: _uRaw := 16#07;   // 段 abc / Segments a b c
8: _uRaw := 16#7F;   // 全七段 / All seven segments
9: _uRaw := 16#6F;   // 段 abcdfg / Segments a b c d f g
ELSE
    _uRaw := 16#00;  // 兜底全灭 / Fallback blanks all
END_CASE

(* 段 3：极性切换 + 单一出口裁决（N4） *)
IF bCommonAnode THEN uSegCode := NOT _uRaw; ELSE uSegCode := _uRaw; END_IF
bValid := TRUE;  FC_DL_SevenSegBcdDecode := TRUE;
END_FUNCTION

(* ---- FC_DL_SevenSegBlankMaskCalc.st ---- *)
(* ============================================================
   DL_Base / FC_DL_SevenSegBlankMaskCalc ｜ v1.0.0 ｜ 2026-11-25
   功能：前导零消隐掩码。uDigitMask 为在位位图（bit i = 第 i+1 位存在），
         uDigits 为有效位数，输出 = 在位位图 ∧ 低 uDigits 位全 1
   边界：uDigits = 0 → 全灭 16#00；uDigits > 8 → 钳到 8 并置码 1（防移位越界）；
         移位量恒 ≤ 7（8 位时改用全 1 常量，禁 SHL 8 位）
   依赖：仅 IEC 61131-3（SHL） ｜ 溯源：DLF-C-SEVENSEG（内部原创线）
   ============================================================ *)
FUNCTION FC_DL_SevenSegBlankMaskCalc : BOOL
VAR_INPUT
    uDigitMask : BYTE;  // 在位位图（bit i = 第 i+1 位存在）[-] / Presence bitmap of the digits
    uDigits    : UINT;  // 有效位数，0 = 无有效位 [位] / Significant digit count
END_VAR
VAR_OUTPUT
    uMask  : BYTE;   // 前导零消隐后允许点亮的位掩码 [-] / Blank mask of allowed digits
    uErrId : UDINT;  // 出口码 0 正常 / 1 有效位数超 8 已钳 [-] / Outlet code
END_VAR
VAR
    _uDigitsUse : UINT;  // 钳定后的有效位数 [位] / Clamped significant digit count
    _uLowOnes   : BYTE;  // 低 n 位全 1 掩码 [-] / Mask with the low n bits set
    _uShiftSrc  : BYTE;  // 移位源（显式 BYTE，禁字面量被推成 DINT）[-] / Explicit BYTE shift source
    _nShift     : INT;   // 归一后移位量（域闸已证 1~7）[位] / Normalized shift amount
END_VAR

(* 段 0：出口预置安全侧（全灭，N3） *)
FC_DL_SevenSegBlankMaskCalc := FALSE;
uMask := 16#00;  uErrId := 0;  _uLowOnes := 16#00;

(* 段 1：位数域闸（0 = 全灭；> 8 钳定并报码） *)
IF uDigits = 0 THEN
    uMask := 16#00;  FC_DL_SevenSegBlankMaskCalc := TRUE;  RETURN;
END_IF
IF uDigits > 8 THEN
    _uDigitsUse := 8;  uErrId := 1;
ELSE
    _uDigitsUse := uDigits;
END_IF

(* 段 2：低 n 位全 1（n = 8 时用全 1 常量，禁 8 位移位；
   移位源与移位量均显式定型：BYTE 源 + INT 量，禁裸字面量被推成 DINT，R48） *)
IF _uDigitsUse >= 8 THEN
    _uLowOnes := 16#FF;
ELSE
    _uShiftSrc := 16#01;                       // 字面量按 BYTE 目标定型
    _nShift    := UINT_TO_INT(_uDigitsUse);    // 域闸已证 1~7，恒 < 位宽 8
    _uLowOnes  := SHL(_uShiftSrc, _nShift) - 16#01;
END_IF

(* 段 3：与在位位图求交（不得点亮硬件不存在的位） + 单一出口裁决（N4） *)
uMask := uDigitMask AND _uLowOnes;
FC_DL_SevenSegBlankMaskCalc := TRUE;
END_FUNCTION

(* ---- FC_DL_SevenSegBlinkPhaseCalc.st ---- *)
(* ============================================================
   DL_Base / FC_DL_SevenSegBlinkPhaseCalc ｜ v1.0.0 ｜ 2026-11-25
   功能：段码闪烁相位判定（毫秒整数域）：rem = tNow MOD tPeriod，
         bOn = (rem < tOn)，fPhase = rem / tPeriod ∈ [0,1)
   边界：tPeriod ≤ 0 → 恒定点亮（bOn=TRUE、fPhase=1.0，N3 先亮最安全）；
         tOn ≤ 0 → 恒定点灭；tOn > tPeriod → 钳到 tPeriod；tNow < 0 按 0；
         MOD 除子已闸非零，无浮点判等（R4）
   依赖：仅 IEC 61131-3（TIME_TO_DINT / DINT_TO_REAL） ｜ 溯源：DLF-C-SEVENSEG
   ============================================================ *)
FUNCTION FC_DL_SevenSegBlinkPhaseCalc : BOOL
VAR_INPUT
    tNow    : TIME;  // 当前时刻（任务时基）[ms] / Current task time base
    tOn     : TIME;  // 一个周期内点亮时长 [ms] / On duration inside one period
    tPeriod : TIME;  // 闪烁周期，> 0 才闪烁 [ms] / Blink period, only a positive value blinks
END_VAR
VAR_OUTPUT
    bOn    : BOOL;  // 本拍应点亮 [-] / Segment should be lit this scan
    fPhase : REAL;  // 周期内相位 [0,1) [-] / Phase inside the period
END_VAR
VAR
    _nNow    : DINT;  // 当前时刻毫秒值 [ms] / Current time in milliseconds
    _nPeriod : DINT;  // 周期毫秒值 [ms] / Period in milliseconds
    _nOn     : DINT;  // 点亮时长毫秒值（已钳定）[ms] / Clamped on duration
    _nRem    : DINT;  // 周期内余量 [ms] / Remainder inside the period
END_VAR

(* 段 0：出口预置安全侧（先亮，无显示熄灭风险） *)
FC_DL_SevenSegBlinkPhaseCalc := FALSE;
bOn := TRUE;  fPhase := 1.0;

(* 段 1：周期域闸（≤ 0 → 恒亮） *)
_nPeriod := TIME_TO_DINT(tPeriod);
IF _nPeriod <= 0 THEN
    bOn := TRUE;  fPhase := 1.0;  FC_DL_SevenSegBlinkPhaseCalc := TRUE;  RETURN;
END_IF

(* 段 2：时刻与点亮时长归一（负时刻按 0；tOn 钳到 [0, tPeriod]） *)
_nNow := TIME_TO_DINT(tNow);
IF _nNow < 0 THEN _nNow := 0; END_IF              // 时刻回绕：不产生负相位
_nOn := TIME_TO_DINT(tOn);
IF _nOn < 0 THEN
    _nOn := 0;
ELSIF _nOn > _nPeriod THEN
    _nOn := _nPeriod;                             // 占空 100%
END_IF

(* 段 3：相位与点亮判据（除子已证 > 0） *)
_nRem := _nNow MOD _nPeriod;
fPhase := DINT_TO_REAL(_nRem) / DINT_TO_REAL(_nPeriod);
IF _nRem < _nOn THEN bOn := TRUE; ELSE bOn := FALSE; END_IF

(* 段 4：相位复检（越 [0,1) 即钳，N4） *)
IF (fPhase <> fPhase) OR (fPhase < 0.0) OR (fPhase >= 1.0) THEN fPhase := 0.0; END_IF
FC_DL_SevenSegBlinkPhaseCalc := TRUE;
END_FUNCTION

(* ---- FC_DL_SevenSegBrightnessPwmCalc.st ---- *)
(* ============================================================
   DL_Base / FC_DL_SevenSegBrightnessPwmCalc ｜ v1.0.0 ｜ 2026-11-25
   功能：亮度 → PWM 占空换算：uDuty = uLevel×255/uFullScale（整数式），
         再按下限保护抬到 uMinDuty 并置 bAtMin（防人眼可辨的熄灭/闪烁）
   边界：uFullScale = 0 → 除零闸，占空 0、bAtMin=TRUE、返回 FALSE（N1）；
         uLevel > uFullScale → 按满占空钳定；中间乘积用 UDINT 承载
         （255×255 = 65025 > USINT），防窄型溢出
   依赖：仅 IEC 61131-3（USINT_TO_UDINT / UDINT_TO_USINT） ｜ 溯源：DLF-C-SEVENSEG
   ============================================================ *)
FUNCTION FC_DL_SevenSegBrightnessPwmCalc : BOOL
VAR_INPUT
    uLevel     : USINT;  // 亮度等级，域 0~uFullScale [级] / Brightness level
    uFullScale : USINT;  // 亮度满量程，域 > 0 [级] / Full scale of the brightness
    uMinDuty   : USINT;  // 占空下限保护 [1/255] / Lower duty clamp
END_VAR
VAR_OUTPUT
    uDuty  : USINT;  // 占空值（255 = 100%）[1/255] / Duty value where 255 is one hundred percent
    bAtMin : BOOL;   // 占空被下限抬升 [-] / Duty raised by the lower clamp
END_VAR
VAR
    _uLevelUse : USINT;  // 钳定后亮度等级 [级] / Clamped brightness level
    _udDuty    : UDINT;  // 占空中间值 [1/255] / Intermediate duty value
END_VAR

(* 段 0：出口预置安全侧（占空 0、标志置位，N1/N3） *)
FC_DL_SevenSegBrightnessPwmCalc := FALSE;
uDuty := 0;  bAtMin := TRUE;

(* 段 1：除零闸（满量程为 0 无定义） *)
IF uFullScale = 0 THEN RETURN; END_IF

(* 段 2：等级钳定（超满量程按满占空，禁窄型溢出） *)
IF uLevel > uFullScale THEN _uLevelUse := uFullScale; ELSE _uLevelUse := uLevel; END_IF

(* 段 3：占空换算（UDINT 承载，除子已证 > 0） *)
_udDuty := USINT_TO_UDINT(_uLevelUse) * 255 / USINT_TO_UDINT(uFullScale);
IF _udDuty > 255 THEN _udDuty := 255; END_IF       // 结构性兜底：比例上界 255

(* 段 4：下限保护（判据在原始占空上，出口单点裁决，N4） *)
IF UDINT_TO_USINT(_udDuty) < uMinDuty THEN
    uDuty := uMinDuty;  bAtMin := TRUE;
ELSE
    uDuty := UDINT_TO_USINT(_udDuty);  bAtMin := FALSE;
END_IF
FC_DL_SevenSegBrightnessPwmCalc := TRUE;
END_FUNCTION

(* ---- FC_DL_SevenSegGhostGuardCalc.st ---- *)
(* ============================================================
   DL_Base / FC_DL_SevenSegGhostGuardCalc ｜ v1.0.0 ｜ 2026-11-25
   功能：鬼影抑制消隐时长：tBlank = 段关断延时 + 位切换时间；强驱动模式再留 50%
         余量（1.5 倍），保证「先关全段 → 换位选 → 点新段」的间隙足够
   边界：任一时长 < 0（TIME 负值）→ bCfgBad=TRUE、tBlank=T#0S（不给不可信时长）；
         tBlank > 5ms（超常规 1ms 位槽上限）→ 钳到 5ms 并置 bCfgBad；
         精度声明：本件以 DINT 毫秒为运算域
   依赖：仅 IEC 61131-3（TIME_TO_DINT / DINT_TO_TIME） ｜ 溯源：DLF-C-SEVENSEG
   ============================================================ *)
FUNCTION FC_DL_SevenSegGhostGuardCalc : BOOL
VAR_INPUT
    tSegOff      : TIME;  // 段关断延时，域 ≥ 0 [ms] / Segment turn off delay
    tDigitSwitch : TIME;  // 位选切换时间，域 ≥ 0 [ms] / Digit select switching time
    bFastMode    : BOOL;  // TRUE=强驱动，留 50% 余量 [-] / TRUE adds fifty percent margin
END_VAR
VAR_OUTPUT
    tBlank  : TIME;  // 计算所得消隐时长 [ms] / Computed blanking duration
    bCfgBad : BOOL;  // 组态非法或时长越上限 [-] / Illegal configuration or above the ceiling
END_VAR
VAR
    _nSeg   : DINT;  // 段关断延时毫秒值 [ms] / Segment turn off delay
    _nBlank : DINT;  // 消隐时长中间值 [ms] / Intermediate blanking duration
END_VAR

(* 段 0：出口预置安全侧（不消隐、标非法） *)
FC_DL_SevenSegGhostGuardCalc := FALSE;
tBlank := T#0S;  bCfgBad := TRUE;

(* 段 1：入参域闸（TIME 负值不可用于时长） *)
_nSeg := TIME_TO_DINT(tSegOff);
IF (_nSeg < 0) OR (TIME_TO_DINT(tDigitSwitch) < 0) THEN RETURN; END_IF

(* 段 2：基础消隐 = 段关断 + 位切换（ms 域相加，无 TIME 溢出路径） *)
_nBlank := _nSeg + TIME_TO_DINT(tDigitSwitch);

(* 段 3：强驱动余量 1.5 倍（整数式 blank + blank/2） *)
IF bFastMode THEN _nBlank := _nBlank + (_nBlank / 2); END_IF

(* 段 4：上限栅（超 5ms 判组态异常并钳定，出口与判据同源，N4） *)
IF _nBlank > 5 THEN
    _nBlank := 5;  bCfgBad := TRUE;
ELSE
    bCfgBad := FALSE;
END_IF
tBlank := DINT_TO_TIME(_nBlank);
FC_DL_SevenSegGhostGuardCalc := TRUE;
END_FUNCTION

(* ---- FC_DL_SevenSegGlyphFontCalc.st ---- *)
(* ============================================================
   DL_Base / FC_DL_SevenSegGlyphFontCalc ｜ v1.0.0 ｜ 2026-11-25
   功能：自定义字形字模查表：段掩码（bit0=a … bit6=g，不含 dp）在标准字形表中
         精确匹配，命中输出槽号 uFontSlot（0~15），未命中置 bMiss
   边界：uSlotCnt = 0 → 无槽可查（bMiss=TRUE、槽号 0）；uSlotCnt > 16 → 钳到
         表容量；数组下标一律 INT 循环索引并夹到本表固定界 0..15（固定长度数组
         故用编译期常量界，LOWER_BOUND/UPPER_BOUND 仅接受变长数组，R17）
   依赖：仅 IEC 61131-3（INT_TO_BYTE） ｜ 溯源：DLF-C-SEVENSEG
   ============================================================ *)
FUNCTION FC_DL_SevenSegGlyphFontCalc : BOOL
VAR_INPUT
    uSegMask : BYTE;  // 段掩码（不含 dp）[-] / Segment mask without the decimal point
    uSlotCnt : UINT;  // 可查字形槽数，域 1~16 [槽] / Number of glyph slots to search
END_VAR
VAR_OUTPUT
    uFontSlot : BYTE;  // 命中的字形槽号 [-] / Matched glyph slot number
    bMiss     : BOOL;  // 未命中任何槽 [-] / No glyph slot matched
END_VAR
VAR
    auFont : ARRAY[0..15] OF BYTE;  // 标准字形表（0~9 与 A~F）[-] / Standard glyph table
    _nCnt  : INT;                   // 钳定后槽数 [槽] / Clamped slot count
    _nIdx  : INT;                   // 循环索引（整数、已夹界）[-] / Bounded loop index
    _bHit  : BOOL;                  // 命中标志 [-] / Match found flag
END_VAR

(* 段 0：出口预置安全侧（槽 0、未命中） *)
FC_DL_SevenSegGlyphFontCalc := FALSE;
uFontSlot := 0;  bMiss := TRUE;  _bHit := FALSE;

(* 段 1：字模表装配（段掩码常量，非码位） *)
auFont[0] := 16#3F;   auFont[1] := 16#06;   auFont[2] := 16#5B;   auFont[3] := 16#4F;
auFont[4] := 16#66;   auFont[5] := 16#6D;   auFont[6] := 16#7D;   auFont[7] := 16#07;
auFont[8] := 16#7F;   auFont[9] := 16#6F;   auFont[10] := 16#77;  auFont[11] := 16#7C;
auFont[12] := 16#39;  auFont[13] := 16#5E;  auFont[14] := 16#79;  auFont[15] := 16#71;

(* 段 2：槽数域闸（0 = 无槽；> 16 钳到表容量） *)
IF uSlotCnt = 0 THEN
    bMiss := TRUE;  FC_DL_SevenSegGlyphFontCalc := TRUE;  RETURN;
END_IF
IF UINT_TO_INT(uSlotCnt) > 15 THEN         // 15 = 固定表上界（auFont[0..15]）
    _nCnt := 16;                              // 钳定到表容量，防越界
ELSE
    _nCnt := UINT_TO_INT(uSlotCnt);
END_IF

(* 段 3：线性查表（索引恒在固定界 0..15 内） *)
FOR _nIdx := 0 TO (_nCnt - 1) DO
    IF (_nIdx >= 0) AND (_nIdx <= 15) THEN
        IF auFont[_nIdx] = uSegMask THEN
            uFontSlot := INT_TO_BYTE(_nIdx);  // 命中：输出槽号
            _bHit := TRUE;
            EXIT;
        END_IF
    END_IF
END_FOR

(* 段 4：单一出口裁决（N4：命中位与槽号同源） *)
bMiss := NOT _bHit;  FC_DL_SevenSegGlyphFontCalc := TRUE;
END_FUNCTION

(* ---- FC_DL_SevenSegHexCodeCalc.st ---- *)
(* ============================================================
   DL_Base / FC_DL_SevenSegHexCodeCalc ｜ v1.0.0 ｜ 2026-11-25
   功能：0~15 十六进制字形段码（A~F 近似字形），段位口径同族（bit0=a … bit6=g）
   边界：uHex > 15 → 全灭 + 码 1；bHexMode=FALSE 且 10~15 → 全灭 + 码 2；
         共阳「全灭」= 16#FF，极性切换在单一出口段完成（N4）；
         16# 常量均为段掩码，非事件码位（R83 不入账）
   依赖：仅 IEC 61131-3（NOT / BYTE_TO_UDINT） ｜ 溯源：DLF-C-SEVENSEG（内部原创线）
   ============================================================ *)
FUNCTION FC_DL_SevenSegHexCodeCalc : BOOL
VAR_INPUT
    uHex         : BYTE;  // 十六进制位值，域 0~15 [-] / Hexadecimal digit, domain zero to fifteen
    bHexMode     : BOOL;  // TRUE=十六进制 / FALSE=BCD 严格校验 [-] / TRUE enables hexadecimal glyphs
    bCommonAnode : BOOL;  // TRUE=共阳低有效 [-] / TRUE for common anode active low
END_VAR
VAR_OUTPUT
    uSegCode : BYTE;   // 七段段码（含极性，不含 dp）[-] / Segment code with polarity
    uErrId   : UDINT;  // 出口码 0 正常 / 1 超 15 / 2 BCD 域外 [-] / Outlet code
END_VAR
VAR
    _uRaw : BYTE;  // 共阴原始段码 [-] / Raw common cathode code
END_VAR

(* 段 0：出口预置安全侧（全灭按极性、码取最严） *)
FC_DL_SevenSegHexCodeCalc := FALSE;
_uRaw := 16#00;  uErrId := 1;
IF bCommonAnode THEN uSegCode := 16#FF; ELSE uSegCode := 16#00; END_IF

(* 段 1：输入域闸与模式闸（BYTE 无符号，单侧判即够） *)
IF BYTE_TO_UDINT(uHex) > 15 THEN RETURN; END_IF
IF (NOT bHexMode) AND (BYTE_TO_UDINT(uHex) > 9) THEN uErrId := 2; RETURN; END_IF

(* 段 2：字形查表（段掩码常量） *)
CASE uHex OF
0:  _uRaw := 16#3F;  // 字形 0 / Glyph zero
1:  _uRaw := 16#06;  // 字形 1 / Glyph one
2:  _uRaw := 16#5B;  // 字形 2 / Glyph two
3:  _uRaw := 16#4F;  // 字形 3 / Glyph three
4:  _uRaw := 16#66;  // 字形 4 / Glyph four
5:  _uRaw := 16#6D;  // 字形 5 / Glyph five
6:  _uRaw := 16#7D;  // 字形 6 / Glyph six
7:  _uRaw := 16#07;  // 字形 7 / Glyph seven
8:  _uRaw := 16#7F;  // 字形 8 / Glyph eight
9:  _uRaw := 16#6F;  // 字形 9 / Glyph nine
10: _uRaw := 16#77;  // 近似字形 A / Approximated glyph A
11: _uRaw := 16#7C;  // 近似字形 b / Approximated glyph b
12: _uRaw := 16#39;  // 近似字形 C / Approximated glyph C
13: _uRaw := 16#5E;  // 近似字形 d / Approximated glyph d
14: _uRaw := 16#79;  // 近似字形 E / Approximated glyph E
15: _uRaw := 16#71;  // 近似字形 F / Approximated glyph F
ELSE
    _uRaw := 16#00;  // 兜底全灭 / Fallback blanks all
END_CASE

(* 段 3：极性切换 + 单一出口裁决（N4） *)
IF bCommonAnode THEN uSegCode := NOT _uRaw; ELSE uSegCode := _uRaw; END_IF
uErrId := 0;  FC_DL_SevenSegHexCodeCalc := TRUE;
END_FUNCTION

(* ---- FC_DL_SevenSegMinusFlagCalc.st ---- *)
(* ============================================================
   DL_Base / FC_DL_SevenSegMinusFlagCalc ｜ v1.0.0 ｜ 2026-11-25
   功能：修饰段叠加 —— 负号段 g(bit6) 与小数点段 dp(bit7) 按位或叠加到字形段码；
         契约对齐 FC_DL_SevenSegBcdDecode：该件头注指名 dp 叠加归本件负责，
         且该件已按 bCommonAnode 输出带极性的段码，本件同口径补极性引脚。
   极性：bCommonAnode=FALSE → 共阴高有效（置位 = 点亮）；TRUE → 共阳低有效。
         实现内部一律先归一到共阴域叠加，再回到调用方口径——禁在共阳（低有效）
         码上直接置位（那会把对应段置 1 即熄灭，表现为「叠加即灭段」）。
   边界：段占用冲突（请求位在原段码中已亮）→ 冲突位不叠加、返回 FALSE
         （签名无独立 BOOL 口，返回值承载 bOverflow 语义，与名称同源以免名实不符）；
         无修饰请求 → 原样透传（极性原样，不做取反）返回 TRUE
   依赖：仅 IEC 61131-3（AND / OR / XOR） ｜ 溯源：DLF-C-SEVENSEG（内部原创线）
   ============================================================ *)
FUNCTION FC_DL_SevenSegMinusFlagCalc : BOOL
VAR_INPUT
    uSegCode      : BYTE;  // 原字形段码（含极性，不含修饰段）[-] / Base glyph code carrying the polarity
    bCommonAnode  : BOOL;  // TRUE=共阳低有效 / FALSE=共阴高有效 [-] / TRUE for common anode wiring
    bMinus        : BOOL;  // 请求叠加负号段 g [-] / Request the minus segment
    bDecimalPoint : BOOL;  // 请求叠加小数点段 dp [-] / Request the decimal point segment
END_VAR
VAR_OUTPUT
    uSegCodeOut : BYTE;  // 叠加后段码（与输入同极性）[-] / Resulting code in the same polarity
END_VAR
VAR
    _uWant : BYTE;  // 请求叠加的修饰段掩码（共阴域高有效）[-] / Requested modifier mask in the common cathode domain
    _uBase : BYTE;  // 极性归一后的共阴高有效段码 [-] / Base code normalized to the common cathode domain
    _uOut  : BYTE;  // 共阴域叠加结果 [-] / Overlaid code in the common cathode domain
END_VAR

(* 段 0：出口预置（空码，N3） *)
FC_DL_SevenSegMinusFlagCalc := TRUE;
uSegCodeOut := 16#00;  _uWant := 16#00;  _uBase := 16#00;  _uOut := 16#00;

(* 段 1：极性归一（共阳低有效取反到共阴高有效域，叠加只在共阴域进行） *)
IF bCommonAnode THEN
    _uBase := uSegCode XOR 16#FF;               // 低有效码逐位取反 → 高有效语义
ELSE
    _uBase := uSegCode;
END_IF

(* 段 1b：组装修饰掩码（g = 16#40，dp = 16#80，共阴域高有效） *)
IF bMinus THEN _uWant := _uWant OR 16#40; END_IF
IF bDecimalPoint THEN _uWant := _uWant OR 16#80; END_IF

(* 段 2：无修饰请求 → 原样透传（极性随原码，不做取反） *)
IF _uWant = 16#00 THEN
    uSegCodeOut := uSegCode;  FC_DL_SevenSegMinusFlagCalc := TRUE;  RETURN;
END_IF

(* 段 3：段占用冲突检测（判据与出口同源：均基于归一后的原始段码） *)
IF (_uBase AND _uWant) <> 16#00 THEN
    uSegCodeOut := uSegCode;                 // 冲突位不重复叠加，保持原码
    FC_DL_SevenSegMinusFlagCalc := FALSE;    // 返回值承载段占用冲突语义
    RETURN;
END_IF

(* 段 4：叠加（共阴域位或，再按调用方口径回送，单一出口裁决 N4） *)
_uOut := _uBase OR _uWant;
IF bCommonAnode THEN
    uSegCodeOut := _uOut XOR 16#FF;          // 回到共阳低有效口径（置 0 = 点亮）
ELSE
    uSegCodeOut := _uOut;
END_IF
FC_DL_SevenSegMinusFlagCalc := TRUE;
END_FUNCTION

(* ---- FC_DL_SevenSegMultiplexPhaseCalc.st ---- *)
(* ============================================================
   DL_Base / FC_DL_SevenSegMultiplexPhaseCalc ｜ v1.0.0 ｜ 2026-11-25
   功能：多路扫描相位解算：每位槽时长 tSlot = tScan / uDigitCnt，
         位索引 uDigitIdx = (tNow MOD tScan) / tSlot（0 基）
   边界：uDigitCnt = 0（位缺失）→ 索引 0、tSlot=T#0S；uDigitCnt > 8 → 钳到 8；
         tScan ≤ 0 → 不做除法（R4 除零闸）；槽时长 < 1ms → 抬到 1ms，
         防位索引恒 0 的隐性命中；全程整数域，无浮点判等
   依赖：仅 IEC 61131-3（TIME_TO_DINT / DINT_TO_TIME） ｜ 溯源：DLF-C-SEVENSEG
   ============================================================ *)
FUNCTION FC_DL_SevenSegMultiplexPhaseCalc : BOOL
VAR_INPUT
    tNow      : TIME;  // 当前时刻（任务时基）[ms] / Current task time base
    uDigitCnt : UINT;  // 扫描位数，域 1~8 [位] / Scanned digit count
    tScan     : TIME;  // 整帧扫描周期，域 > 0 [ms] / Frame scan period
END_VAR
VAR_OUTPUT
    uDigitIdx : UINT;  // 当前位索引（0 基）[-] / Current digit index starting at zero
    tSlot     : TIME;  // 每位保持时间 [ms] / Hold time of one digit slot
END_VAR
VAR
    _nScanMs : DINT;  // 帧周期毫秒值 [ms] / Frame period in milliseconds
    _nCnt    : DINT;  // 钳定后位数 [位] / Clamped digit count
    _nSlotMs : DINT;  // 每槽毫秒值 [ms] / Slot duration in milliseconds
    _nIdx    : DINT;  // 位索引中间值 [-] / Intermediate digit index
END_VAR

(* 段 0：出口预置安全侧（索引 0、槽时长 0） *)
FC_DL_SevenSegMultiplexPhaseCalc := FALSE;
uDigitIdx := 0;  tSlot := T#0S;

(* 段 1：位数域闸（0 = 无位可扫；> 8 钳定） *)
IF uDigitCnt = 0 THEN RETURN; END_IF
_nCnt := UINT_TO_DINT(uDigitCnt);
IF _nCnt > 8 THEN _nCnt := 8; END_IF

(* 段 2：帧周期域闸（≤ 0 不做除法） *)
_nScanMs := TIME_TO_DINT(tScan);
IF _nScanMs <= 0 THEN RETURN; END_IF

(* 段 3：槽时长（除子 ∈ 1..8，除零结构不可达） *)
_nSlotMs := _nScanMs / _nCnt;
IF _nSlotMs < 1 THEN _nSlotMs := 1; END_IF        // 抬到 1ms，防索引恒 0
tSlot := DINT_TO_TIME(_nSlotMs);

(* 段 4：帧内余量与位索引（钳到 0..cnt−1，防越界） *)
_nIdx := TIME_TO_DINT(tNow);
IF _nIdx < 0 THEN _nIdx := 0; END_IF              // 时刻回绕：按 0 处理
_nIdx := (_nIdx MOD _nScanMs) / _nSlotMs;         // 两除子均已证 > 0
IF _nIdx >= _nCnt THEN _nIdx := _nCnt - 1; END_IF
IF _nIdx < 0 THEN _nIdx := 0; END_IF
uDigitIdx := DINT_TO_UINT(_nIdx);

(* 段 5：单一出口裁决（N4） *)
FC_DL_SevenSegMultiplexPhaseCalc := TRUE;
END_FUNCTION

(* ---- FC_DL_ShiftArithEx.st ---- *)
(*
  ==================================================================
  组件名 Component  : FC_DL_ShiftArithEx
  分类   Category   : DL_Base
  前缀   Naming     : FC_DL_ ｜ b/n/u/f/t/e/st 类型前缀制（R265）
  码位   Code ID    : 16#0001_064B（信息级）｜ 16#0001_064C（信息级）
  版本   Version    : 1.0.0
  复杂度 Complexity  : 中
  功能   Purpose    : DINT 算术右移（符号位扩展右移）：IEC 标准只有逻辑 SHR，本件补
                      算术语义，移位量越域按语义钳位并以 bSat 提示。
  开源溯源 Origin    : IEC 61131-3 标准语义的道莅防御性实现（clean-room，无第三方代码行）
  许可证 License    : MIT
  参考   Reference  : IEC 61131-3:2013 §6.6.3 位串移位函数 SHR 的语义与实参域
  平台   Platform   : 纯 IEC 61131-3（SHR / OR / 类型转换），CODESYS / TwinCAT 3 / InoProShop 通用
  依赖   Depends    : 仅 Standard.library（SHR 属标准位串函数）
  分工声明 Split     : FC_DL_ShrEx（DWORD 逻辑右移）与 FC_DL_ShrLwordEx（LWORD 逻辑
                      右移）为逻辑右移属主，本件不重复其职责；IEC 标准无算术右移原语，
                      故本件仅补符号扩展语义（R216 双向互引）。
  归属 Ownership     : 本件无 TYPE 声明；常量表 DL_SAR_MASK 为本文件私有常量。
  ------------------------------------------------------------------
  边界 Boundary     :
                      一 移位量归一（R48）：nShift ≥ 32 时不调用 SHR，直接走「全符号位
                         填充」常量路径，杜绝 SHL/SHR(x, 32) 的未定义行为；
                      二 高位掩码用 32 项预计算常量表，禁运行时 SHL(x, 32)；
                         掩码仅在符号位为 1 时参与 OR，否则会把非负结果污染成负数；
                      三 nShift ≤ 0 原值返回（0 移位不改值）；nShift < 0 反向移位非法，
                         钳 0 并置 bSat + 信息码，禁静默反向移位；
                      四 纯函数：无记忆量、无定时器、无边沿实例，每调用重算。
  错误码 Codes      :
    16#0001_064B【信息级】移位量为负已钳 0（反向移位非法，结果等于原值）
    16#0001_064C【信息级】移位量 ≥ 32 已按符号位全填充饱和（负数得 -1，非负得 0）
  码位反证 Note     :
    064B 与 064C 不可合并：两者 bSat 同为 TRUE，但「原值返回」与「全符号填充」是
    两个相反的语义分支，合并后现场无法由 diOut 与 bSat 唯一还原是哪种越域（R90）。
  验收 Acceptance   :
    算法已证（脚本）：未跑 ｜ 编译器已证（三平台）：未跑
    V1 -8 >> 1 → -4；V2 -1 >> 5 → -1（全 1 保持）；V3 8 >> 31 → 0
    V4 8 >> 32 → 0 且 bSat = TRUE、码 064C
    V5 -8 >> 32 → -1 且 bSat = TRUE（符号填充）
    V6 x >> 0 → x 精确、bSat = FALSE、无码
    V7 x >> -1 → x 且 bSat = TRUE、码 064B（越域钳 0）
    V8 MIN >> 1 → -1073741824（符号保持）
  修订记录 Revision  :
    2026-11-21  v1.0.0  R62 首版（批 1 · 序号 3）
  ==================================================================
*)
FUNCTION FC_DL_ShiftArithEx : BOOL
VAR_INPUT
    diIn   : DINT; // 待移位值 [−]，完整 DINT 域 / the value to shift over the full DINT domain
    nShift : DINT; // 移位位数 [位]，合法域 1..31，0 原值、负值钳 0、≥32 饱和 / the shift amount in bits, valid one to thirty one
END_VAR
VAR_OUTPUT
    diOut  : DINT;  // 算术右移结果 [−] / the arithmetic shift result
    bSat   : BOOL;  // 移位量越域已被钳（含负值与 ≥32）[-] / the shift amount was out of domain and clamped
    eErr   : UDINT; // 错误码，0 = 正常 / the error code, zero is ok
    bError : BOOL;  // 故障标志（本件只有信息级码，恒 FALSE，保留引脚供族内统一）/ the fault flag, always false here since only informational codes exist
END_VAR
VAR
    udwWork : DWORD := 16#0000_0000; // 逻辑右移工作寄存器 [位] / the logical shift working register in bits
    nUse    : DINT := 0;             // 归一后的移位量 [位] / the normalized shift amount in bits
END_VAR  // R64 结构补齐：VAR 段缺失的 END_VAR（门禁机械修复）
VAR CONSTANT
    DL_SAR_ZERO : DINT := 0;         // 零常量 [位] / the zero constant
    DL_SAR_BITS : DINT := 32;        // DINT 容器位宽 [位] / the DINT container width in bits
    DL_SAR_NEG1 : DINT := -1;        // 全 1 常量（负数饱和填充值）[−] / the all ones constant used as the negative saturation fill
    DL_SAR_MASK : ARRAY[0..31] OF DWORD := // 高位掩码表（第 k 项 = 高 k 位置 1，k = 0 为零），预计算禁运行时 SHL(x,32) [位] / the precomputed high side mask table, k bits set from the top
    [
        16#0000_0000, // k = 0：不移位，无高位 / k equals zero, no high bits at all
        16#8000_0000, // k = 1：最高 1 位 / the top single bit
        16#C000_0000, // k = 2 / two top bits
        16#E000_0000, // k = 3 / three top bits
        16#F000_0000, // k = 4 / four top bits
        16#F800_0000, // k = 5 / five top bits
        16#FC00_0000, // k = 6 / six top bits
        16#FE00_0000, // k = 7 / seven top bits
        16#FF00_0000, // k = 8 / eight top bits
        16#FF80_0000, // k = 9 / nine top bits
        16#FFC0_0000, // k = 10 / ten top bits
        16#FFE0_0000, // k = 11 / eleven top bits
        16#FFF0_0000, // k = 12 / twelve top bits
        16#FFF8_0000, // k = 13 / thirteen top bits
        16#FFFC_0000, // k = 14 / fourteen top bits
        16#FFFE_0000, // k = 15 / fifteen top bits
        16#FFFF_0000, // k = 16：高半字 / the whole high half word
        16#FFFF_8000, // k = 17 / seventeen top bits
        16#FFFF_C000, // k = 18 / eighteen top bits
        16#FFFF_E000, // k = 19 / nineteen top bits
        16#FFFF_F000, // k = 20 / twenty top bits
        16#FFFF_F800, // k = 21 / twenty one top bits
        16#FFFF_FC00, // k = 22 / twenty two top bits
        16#FFFF_FE00, // k = 23 / twenty three top bits
        16#FFFF_FF00, // k = 24 / twenty four top bits
        16#FFFF_FF80, // k = 25 / twenty five top bits
        16#FFFF_FFC0, // k = 26 / twenty six top bits
        16#FFFF_FFE0, // k = 27 / twenty seven top bits
        16#FFFF_FFF0, // k = 28 / twenty eight top bits
        16#FFFF_FFF8, // k = 29 / twenty nine top bits
        16#FFFF_FFFC, // k = 30 / thirty top bits
        16#FFFF_FFFE  // k = 31 / thirty one top bits
    ];
END_VAR

// 段 1｜返回值与全部出口预置安全值（R45 四段式第一段）/ segment 1, preset every outlet to its safe value
FC_DL_ShiftArithEx := FALSE; // 返回值预置假 / preset the return false
diOut := DL_SAR_ZERO; // 结果预置零 [−] / preset the result zero
bSat := FALSE; // 越域标志预置假 / preset the saturation flag false
eErr := 16#0000_0000; // 错误码预置正常 / preset the code to ok
bError := FALSE; // 故障标志预置假（本件无故障级码）/ preset the fault flag false, no fault level code exists here
udwWork := 16#0000_0000; // 工作寄存器清零 [位] / clear the working register
nUse := DL_SAR_ZERO; // 归一移位量清零 [位] / clear the normalized shift amount

// 段 2｜nShift ≤ 0：0 移位原值返回；负值反向移位非法，钳 0 并提示（边界三）/ segment 2, the non positive shift amount branch
IF nShift < DL_SAR_ZERO THEN // 反向移位非法 / a reverse shift is illegal
    bSat := TRUE; // 置越域标志 / raise the out of domain flag
    eErr := 16#0001_064B; // 信息级：移位量为负已钳 0 / informational, a negative amount is clamped to zero
    diOut := diIn; // 钳 0 后等于原值 [−] / with zero shift the result is the original value
    FC_DL_ShiftArithEx := TRUE; // 信息级不阻断，返回成功 / an informational code does not block, return success
    RETURN; // 早退 / early return
END_IF
IF nShift = DL_SAR_ZERO THEN // 零移位：不改值且无任何提示 / a zero shift changes nothing and raises nothing
    diOut := diIn; // 原值直出 [−] / pass the original value through
    FC_DL_ShiftArithEx := TRUE; // 返回成功 / return success
    RETURN; // 早退 / early return
END_IF

// 段 3｜nShift ≥ 32：不调用 SHR，直接按符号位全填充（边界一，禁 SHL/SHR(x,32)）/ segment 3, the at or above container width branch
IF nShift >= DL_SAR_BITS THEN // 移位量达到或超过容器位宽 / the amount reached or exceeded the container width
    bSat := TRUE; // 置越域标志 / raise the out of domain flag
    eErr := 16#0001_064C; // 信息级：移位量 ≥ 32 已按符号位全填充 / informational, the amount at or above thirty two fills with the sign bit
    IF diIn < DL_SAR_ZERO THEN // 负数：全 1 填充 / a negative value fills with all ones
        diOut := DL_SAR_NEG1; // 结果为 -1 [−] / the result is minus one
    ELSE // 非负数：全 0 填充 / a non negative value fills with zeros
        diOut := DL_SAR_ZERO; // 结果为 0 [−] / the result is zero
    END_IF
    FC_DL_ShiftArithEx := TRUE; // 返回成功 / return success
    RETURN; // 早退 / early return
END_IF

// 段 4｜1 ≤ nShift ≤ 31：逻辑右移 + 符号位为 1 时 OR 高位掩码（边界二）/ segment 4, the normal arithmetic shift by mask
nUse := nShift; // 域内移位量接管（已证 1..31）[位] / take the in-domain amount, proven one to thirty one
udwWork := SHR(DINT_TO_DWORD(diIn), nUse); // 逻辑右移（高位补 0）[位] / the logical shift with zeros shifted in
IF diIn < DL_SAR_ZERO THEN // 符号位为 1 才需补 1（非负数 OR 掩码会污染成负数）/ fill only for a set sign bit, otherwise the mask would turn the result negative
    udwWork := udwWork OR DL_SAR_MASK[nUse]; // 补入高 nUse 个 1 [位] / fill the top amount of ones
END_IF
diOut := DWORD_TO_DINT(udwWork); // 位型还原为有符号结果 [−] / reinterpret the bit pattern as a signed result

// 段 5｜统一出口（信息级未触发，码保持 0）/ segment 5, the unified outlet without any event
bSat := FALSE; // 正常路径明确落假（越域分支已早退）/ the normal path explicitly falls to false, the out of domain branches returned earlier
FC_DL_ShiftArithEx := TRUE; // 返回成功 / return success
END_FUNCTION

(* ---- FC_DL_ShlEx.st ---- *)
(*==============================================================================
 * 组件名称 (Component)  : FC_DL_ShlEx
 * 所属子库 (Sublibrary) : DL_Base
 * 当前版本 (Version)    : 1.0.0
 * 兼容性   (Platform)   : CODESYS 3.5 / TwinCAT 3 / 汇川 InoProShop / Machine Expert
 *                         仅依赖 Standard.library 的 SHL 内建函数，无厂商方言
 * 功能一句话 (Summary)  : 左移防御包装：移位量钳位归一 + 超宽结果零值显式化。
 * 功能描述 (Function)   : 对被移位位串按移位量 nN 左移。nN ≥ 32（位宽）时走常量
 *                         路径直接置 0（严禁 SHL(x, n) 中 n ≥ 位宽的未定义/平台
 *                         歧义行为，R10 BitFieldExtract 先例口径）；nN < 32 才
 *                         委托内建 SHL。纯函数，无内部状态、无跨周期残留。
 * 溯源     (Origin)     : IEC 61131-3 标准语义的道莅防御性实现
 *                         （接口语义由 IEC 61131-3 定义，clean-room 重写，
 *                         参考公开标准条款）
 * 支持位宽 (Width Note) : 本件按 DWORD（32 位）主类型实现，仅支持 32 位位串；
 *                         BYTE / WORD 调用方先显式转换到 DWORD 后调用，再按需
 *                         截回原位宽（头注释显式声明，不做 ANY_BIT 泛型）。
 * 类型裁定 (Type Note)  : 码位段 16#0001_xxxx 为全库共享 32 位段，WORD 容量不足，
 *                         故 uDiag 采用 UDINT 承载（与库内 uErrorId : UDINT 惯例一致）
 * 依赖     (Depends)    : 无 DL_ 内部依赖；Standard.library: SHL
 * 红线自检 (Redline)    : R1 ✓ 零全局变量与外部变量引用 ｜ R2 ✓ 零物理 IO 地址直写
 *                         R3 ✓ 纯 IEC 61131-3 ｜ R4 ✓ 移位量钳位（nN ≥ 32 走常量
 *                         路径）｜ R5 ✓ 全变量中英双语同行注释 ｜ R6 N/A（纯函数，
 *                         无 CASE/ENUM 状态机，按批 1 口径标 N/A）
 *                         R7 N/A（FC 为纯函数，无实例调用，头注释显式说明）
 * 防御行为声明 (Defense): ① nN ≥ 32 时结果直接置 16#0000_0000 并置信息码
 *                           16#0001_0156，不调内建 SHL（部分平台移位量 ≥ 位宽
 *                           属未定义行为或结果歧义，本库统一为「超宽置 0」）；
 *                         ② nN 为 USINT 类型天然非负，nN < 0 不可能发生，
 *                           无负移位量防御分支（类型系统层面保证）；
 *                         ③ 32（位宽）提为只读常量，禁魔法数。
 * 修订历史 (Revision)   :
 *   2026-11-16  v1.0.0  首版入库（R14 批 3 · T0 快车道）
 *============================================================================*)
FUNCTION FC_DL_ShlEx : DWORD
VAR_INPUT
    uIn : DWORD;   // 被移位位串 [位] / Bit string to be shifted
    nN  : USINT;   // 移位量 [bit]，USINT 天然非负 / Shift amount [bit], USINT is non-negative by type
END_VAR
VAR_OUTPUT
    uDiag : UDINT; // 诊断字，16#0001_0156=移位量超宽结果置 0，0=无事件 / Diag word, 16#0001_0156=oversized shift yields zero, 0=no event
END_VAR
VAR CONSTANT
    DL_SH_WIDTH : USINT := 32;  // 位宽常量 [bit]，与 DWORD 位宽一致 / Width constant [bit], matches the DWORD width
END_VAR

(*------------------------------------------------------------------------------
 * 段 1｜输出与诊断预置：先归零，任何路径都不会留下脏诊断
 *      Pre-set the output and diag so no path ever leaves a stale diag
 *-----------------------------------------------------------------------------*)
FC_DL_ShlEx := 16#0000_0000;   // 返回值预置全零 [位串] / Preset return value to all zero
uDiag       := 16#0000_0000;   // 诊断字预置无事件 / Preset diag word to no event

(*------------------------------------------------------------------------------
 * 段 2｜移位量闸门（边界 B1）：nN ≥ 位宽走常量路径直接置 0，不调内建
 *      Shift-amount gate (B1): nN greater or equal to the width takes the
 *      constant path yielding zero, the built-in SHL is never called
 *      严禁把 nN = 32 送进 SHL —— 部分编译器对该移位量属未定义行为
 *      Never feed nN = 32 into SHL, undefined behaviour on some compilers
 *-----------------------------------------------------------------------------*)
IF nN >= DL_SH_WIDTH THEN
    FC_DL_ShlEx := 16#0000_0000;   // 超宽常量路径：结果置 0 [位串] / Oversized constant path: result is zero
    uDiag       := 16#0001_0156;   // 信息码：移位量超宽，结果已置 0 / Informational: oversized shift, result set to zero
ELSE
    FC_DL_ShlEx := SHL(uIn, nN);   // 域内委托内建 SHL，移位量 0 到 31 安全 [位串] / In-domain delegate to built-in SHL, shift amount 0 to 31 is safe
END_IF
END_FUNCTION

(* ---- FC_DL_ShlLwordEx.st ---- *)
(*
    FC_DL_ShlLwordEx —— LWORD 左移（超宽置零）
    ------------------------------------------------------------------
    分类      : DL_Base / BitString
    前缀      : FC_DL_
    版本      : 1.0.0
    溯源      : IEC 61131-3 标准语义的道莅防御性实现
                （接口语义由 IEC 61131-3 定义，内部委托平台内建 SHL，
                  外围统一错误码 / 钳位 / 双语文档；clean-room 重写，
                  未复制任何闭源厂商源码，参考实现仅限 MIT/Apache 许可）
    平台      : 纯 IEC 61131-3，CODESYS / TwinCAT / InoProShop 通用
    作者      : 道莅代码库 · PLC编程专家（R17）
    ------------------------------------------------------------------
    功能说明  : LWORD 位串左移防御包装：移位量 nN 大于等于 64（位宽）时走常量路径直接输出全零，
                并置信息级 16#0001_0233，严禁把 nN ≥ 64 送进内建 SHL
                （部分编译器对该移位量属未定义行为或结果歧义，与 R14 FC_DL_ShlEx 的 32 位口径同源）；
                nN < 64 时委托平台内建 SHL，不重实现移位内核；
                nN 为 USINT 类型天然非负，负移位量结构性不可能（无负值防御分支）；
                位宽 64 提为只读常量，禁魔法数；
                钳位方向：移位量超宽按「结果置 0」处理（不做移位量截断，截断会静默改变语义）。
    错误码    : 16#0001_0233 移位量 ≥ 64（位宽），结果已置全零——信息级，正常防御
                16#0001_0234 预留禁用（信息级，不得挪用）
                16#0001_02F7 预留禁用（故障级，不得挪用）
                16#0001_02F8 预留禁用（故障级，不得挪用）
                16#0001_02F9 预留禁用（故障级，不得挪用）
    状态机    : R6 标注 N/A —— 本组件为纯函数无顺序状态机，无 CASE 可写，非法状态不可能出现，故以本节说明替代 ELSE 兜底
    修订记录  : 2026-11-16 v1.0.0 首次入库（R17）
*)
FUNCTION FC_DL_ShlLwordEx : LWORD
VAR_INPUT
    uIn : LWORD; // 被移位位串 [位] / bit string to be shifted [bit]
    nN  : USINT; // 移位量 [bit]，USINT 天然非负，范围 0~255 / shift amount [bit], USINT is non-negative by type, range 0..255
END_VAR
VAR_OUTPUT
    eErr   : UDINT; // 错误码，0=正常 / error id, 0=ok
    bError : BOOL;  // 是否出错，eErr 非 0 时为 TRUE / error flag, TRUE when eErr is nonzero
    bValid : BOOL;  // 输出是否有效可用 / output valid flag
END_VAR
VAR CONSTANT
    DL_LW_WIDTH : USINT := 64;                        // LWORD 位宽常量 [bit] / LWORD width constant [bit]
    DL_LW_ZERO  : LWORD := 16#0000_0000_0000_0000;     // 超宽移位结果零值 [位串] / zero result of an oversized shift [bit string]
END_VAR

// 段 1｜输出与错误状态预置 / segment 1, preset output and error status
FC_DL_ShlLwordEx := DL_LW_ZERO; // 输出预置全零，任何路径不留脏值 [位串] / preset output to all zeros, no stale value on any path [bit string]
eErr   := 0;     // 预置无错误 / preset no error
bError := FALSE; // 预置无故障（本件无故障级路径） / preset no fault, no fault-level path here
bValid := FALSE; // 预置输出无效，通过移位量闸门后置位 / preset invalid, set TRUE after the shift-amount gate

// 段 2｜移位量闸门（超宽走常量路径，不调内建） / segment 2, shift amount gate (oversized takes the constant path, built-in not called)
IF nN >= DL_LW_WIDTH THEN // 移位量不小于位宽一律走常量路径，绝不送入内建 SHL [bit] / shift amounts not below the width always take the constant path and never reach built-in SHL [bit]
    FC_DL_ShlLwordEx := DL_LW_ZERO; // 结果置全零（不做移位量截断，截断会静默改变语义） [位串] / result set to all zeros, no shift-amount truncation which would silently change semantics [bit string]
    eErr := 16#0001_0233;           // 信息级：超宽移位已置零，正常防御 / info level: oversized shift zeroed, normal defence
    bError := FALSE;                // 信息级不置故障 / info level never raises fault
    bValid := TRUE;                 // 零结果本身有效可用 / the zero result itself is valid
    RETURN;                         // 常量路径即出口，内建 SHL 不被调用 / the constant path is the exit, built-in SHL is not called
END_IF

// 段 3｜域内委托移位（末段） / segment 3, in-domain delegated shift (final)
FC_DL_ShlLwordEx := SHL(uIn, nN); // 域内委托平台内建 SHL，不重实现移位内核 [位串] / in-domain delegate to built-in SHL, shift kernel not re-implemented [bit string]
eErr   := 0;     // 域内无错误 / in-domain, no error
bError := FALSE; // 信息级不置故障 / info level never raises fault
bValid := TRUE;  // 域内输出有效可用 / in-domain output is valid
END_FUNCTION

(* ---- FC_DL_ShrEx.st ---- *)
(*==============================================================================
 * 组件名称 (Component)  : FC_DL_ShrEx
 * 所属子库 (Sublibrary) : DL_Base
 * 当前版本 (Version)    : 1.0.0
 * 兼容性   (Platform)   : CODESYS 3.5 / TwinCAT 3 / 汇川 InoProShop / Machine Expert
 *                         仅依赖 Standard.library 的 SHR 内建函数，无厂商方言
 * 功能一句话 (Summary)  : 右移防御包装：移位量钳位归一 + 超宽结果零值显式化。
 * 功能描述 (Function)   : 对被移位位串按移位量 nN 右移（逻辑右移，高位补 0）。
 *                         nN ≥ 32（位宽）时走常量路径直接置 0（严禁 SHR(x, n)
 *                         中 n ≥ 位宽的未定义/平台歧义行为，R10 BitFieldExtract
 *                         先例口径）；nN < 32 才委托内建 SHR。纯函数，无内部
 *                         状态、无跨周期残留。
 * 溯源     (Origin)     : IEC 61131-3 标准语义的道莅防御性实现
 *                         （接口语义由 IEC 61131-3 定义，clean-room 重写，
 *                         参考公开标准条款）
 * 支持位宽 (Width Note) : 本件按 DWORD（32 位）主类型实现，仅支持 32 位位串；
 *                         BYTE / WORD 调用方先显式转换到 DWORD 后调用，再按需
 *                         截回原位宽（头注释显式声明，不做 ANY_BIT 泛型）。
 * 类型裁定 (Type Note)  : 码位段 16#0001_xxxx 为全库共享 32 位段，WORD 容量不足，
 *                         故 uDiag 采用 UDINT 承载（与库内 uErrorId : UDINT 惯例一致）
 * 依赖     (Depends)    : 无 DL_ 内部依赖；Standard.library: SHR
 * 红线自检 (Redline)    : R1 ✓ 零全局变量与外部变量引用 ｜ R2 ✓ 零物理 IO 地址直写
 *                         R3 ✓ 纯 IEC 61131-3 ｜ R4 ✓ 移位量钳位（nN ≥ 32 走常量
 *                         路径）｜ R5 ✓ 全变量中英双语同行注释 ｜ R6 N/A（纯函数，
 *                         无 CASE/ENUM 状态机，按批 1 口径标 N/A）
 *                         R7 N/A（FC 为纯函数，无实例调用，头注释显式说明）
 * 防御行为声明 (Defense): ① nN ≥ 32 时结果直接置 16#0000_0000 并置信息码
 *                           16#0001_0157，不调内建 SHR（部分平台移位量 ≥ 位宽
 *                           属未定义行为或结果歧义，本库统一为「超宽置 0」）；
 *                         ② nN 为 USINT 类型天然非负，nN < 0 不可能发生，
 *                           无负移位量防御分支（类型系统层面保证）；
 *                         ③ 32（位宽）提为只读常量，禁魔法数。
 * 修订历史 (Revision)   :
 *   2026-11-16  v1.0.0  首版入库（R14 批 3 · T0 快车道）
 *============================================================================*)
FUNCTION FC_DL_ShrEx : DWORD
VAR_INPUT
    uIn : DWORD;   // 被移位位串 [位] / Bit string to be shifted
    nN  : USINT;   // 移位量 [bit]，USINT 天然非负 / Shift amount [bit], USINT is non-negative by type
END_VAR
VAR_OUTPUT
    uDiag : UDINT; // 诊断字，16#0001_0157=移位量超宽结果置 0，0=无事件 / Diag word, 16#0001_0157=oversized shift yields zero, 0=no event
END_VAR
VAR CONSTANT
    DL_SR_WIDTH : USINT := 32;  // 位宽常量 [bit]，与 DWORD 位宽一致 / Width constant [bit], matches the DWORD width
END_VAR

(*------------------------------------------------------------------------------
 * 段 1｜输出与诊断预置：先归零，任何路径都不会留下脏诊断
 *      Pre-set the output and diag so no path ever leaves a stale diag
 *-----------------------------------------------------------------------------*)
FC_DL_ShrEx := 16#0000_0000;   // 返回值预置全零 [位串] / Preset return value to all zero
uDiag       := 16#0000_0000;   // 诊断字预置无事件 / Preset diag word to no event

(*------------------------------------------------------------------------------
 * 段 2｜移位量闸门（边界 B1）：nN ≥ 位宽走常量路径直接置 0，不调内建
 *      Shift-amount gate (B1): nN greater or equal to the width takes the
 *      constant path yielding zero, the built-in SHR is never called
 *      严禁把 nN = 32 送进 SHR —— 部分编译器对该移位量属未定义行为
 *      Never feed nN = 32 into SHR, undefined behaviour on some compilers
 *-----------------------------------------------------------------------------*)
IF nN >= DL_SR_WIDTH THEN
    FC_DL_ShrEx := 16#0000_0000;   // 超宽常量路径：结果置 0 [位串] / Oversized constant path: result is zero
    uDiag       := 16#0001_0157;   // 信息码：移位量超宽，结果已置 0 / Informational: oversized shift, result set to zero
ELSE
    FC_DL_ShrEx := SHR(uIn, nN);   // 域内委托内建 SHR，移位量 0 到 31 安全 [位串] / In-domain delegate to built-in SHR, shift amount 0 to 31 is safe
END_IF
END_FUNCTION

(* ---- FC_DL_ShrLwordEx.st ---- *)
(*
    FC_DL_ShrLwordEx —— LWORD 逻辑右移（超宽置零）
    ------------------------------------------------------------------
    分类      : DL_Base / BitString
    前缀      : FC_DL_
    版本      : 1.0.0
    溯源      : IEC 61131-3 标准语义的道莅防御性实现
                （接口语义由 IEC 61131-3 定义，内部委托平台内建 SHR，
                  外围统一错误码 / 钳位 / 双语文档；clean-room 重写，
                  未复制任何闭源厂商源码，参考实现仅限 MIT/Apache 许可）
    平台      : 纯 IEC 61131-3，CODESYS / TwinCAT / InoProShop 通用
    作者      : 道莅代码库 · PLC编程专家（R17）
    ------------------------------------------------------------------
    功能说明  : LWORD 位串逻辑右移防御包装：移位量 nN 大于等于 64（位宽）时走常量路径直接输出全零，
                并置信息级 16#0001_0232，严禁把 nN ≥ 64 送进内建 SHR；
                nN < 64 时委托平台内建 SHR，不重实现移位内核；
                LWORD 为无符号位串，逻辑右移与算术右移等价，本件不做符号位扩展
                （若调用方需要符号语义，请先用显式类型转换，不得在本件内隐式判断）；
                nN 为 USINT 类型天然非负，负移位量结构性不可能；
                钳位方向：移位量超宽按「结果置 0」处理。
    错误码    : 16#0001_0232 移位量 ≥ 64（位宽），结果已置全零——信息级，正常防御
                16#0001_0209 预留禁用（信息级，不得挪用）
                16#0001_02FA 预留禁用（故障级，不得挪用）
                16#0001_02FB 预留禁用（故障级，不得挪用）
                16#0001_02FC 预留禁用（故障级，不得挪用）
    状态机    : R6 标注 N/A —— 本组件为纯函数无顺序状态机，无 CASE 可写，非法状态不可能出现，故以本节说明替代 ELSE 兜底
    修订记录  : 2026-11-16 v1.0.0 首次入库（R17）
*)
FUNCTION FC_DL_ShrLwordEx : LWORD
VAR_INPUT
    uIn : LWORD; // 被移位位串（无符号位串，无符号位扩展语义） [位] / bit string to be shifted, unsigned, no sign extension [bit]
    nN  : USINT; // 移位量 [bit]，USINT 天然非负，范围 0~255 / shift amount [bit], USINT is non-negative by type, range 0..255
END_VAR
VAR_OUTPUT
    eErr   : UDINT; // 错误码，0=正常 / error id, 0=ok
    bError : BOOL;  // 是否出错，eErr 非 0 时为 TRUE / error flag, TRUE when eErr is nonzero
    bValid : BOOL;  // 输出是否有效可用 / output valid flag
END_VAR
VAR CONSTANT
    DL_LW_WIDTH : USINT := 64;                        // LWORD 位宽常量 [bit] / LWORD width constant [bit]
    DL_LW_ZERO  : LWORD := 16#0000_0000_0000_0000;     // 超宽移位结果零值 [位串] / zero result of an oversized shift [bit string]
END_VAR

// 段 1｜输出与错误状态预置 / segment 1, preset output and error status
FC_DL_ShrLwordEx := DL_LW_ZERO; // 输出预置全零，任何路径不留脏值 [位串] / preset output to all zeros, no stale value on any path [bit string]
eErr   := 0;     // 预置无错误 / preset no error
bError := FALSE; // 预置无故障（本件无故障级路径） / preset no fault, no fault-level path here
bValid := FALSE; // 预置输出无效，通过移位量闸门后置位 / preset invalid, set TRUE after the shift-amount gate

// 段 2｜移位量闸门（超宽走常量路径，不调内建） / segment 2, shift amount gate (oversized takes the constant path, built-in not called)
IF nN >= DL_LW_WIDTH THEN // 移位量不小于位宽一律走常量路径，绝不送入内建 SHR [bit] / shift amounts not below the width always take the constant path and never reach built-in SHR [bit]
    FC_DL_ShrLwordEx := DL_LW_ZERO; // 结果置全零（无符号位串逻辑右移后高位全补 0） [位串] / result set to all zeros, logical right shift of an unsigned string fills zeros [bit string]
    eErr := 16#0001_0232;           // 信息级：超宽移位已置零，正常防御 / info level: oversized shift zeroed, normal defence
    bError := FALSE;                // 信息级不置故障 / info level never raises fault
    bValid := TRUE;                 // 零结果本身有效可用 / the zero result itself is valid
    RETURN;                         // 常量路径即出口，内建 SHR 不被调用 / the constant path is the exit, built-in SHR is not called
END_IF

// 段 3｜域内委托移位（末段） / segment 3, in-domain delegated shift (final)
FC_DL_ShrLwordEx := SHR(uIn, nN); // 域内委托平台内建 SHR，不重实现移位内核 [位串] / in-domain delegate to built-in SHR, shift kernel not re-implemented [bit string]
eErr   := 0;     // 域内无错误 / in-domain, no error
bError := FALSE; // 信息级不置故障 / info level never raises fault
bValid := TRUE;  // 域内输出有效可用 / in-domain output is valid
END_FUNCTION

(* ---- FC_DL_SignExtendEx.st ---- *)
(*
  ==================================================================
  组件名 Component  : FC_DL_SignExtendEx
  分类   Category   : DL_Base
  前缀   Naming     : FC_DL_ ｜ b/n/u/f/t/e/st 类型前缀制（R265）
  码位   Code ID    : 16#0001_064D（故障级）
  版本   Version    : 1.0.0
  复杂度 Complexity  : 中
  功能   Purpose    : 取 DINT 的低 nWidth 位，按 bSigned 选择符号扩展或零扩展，结果落 DINT。
  开源溯源 Origin    : IEC 61131-3 标准语义的道莅防御性实现（clean-room，无第三方代码行）
  许可证 License    : MIT
  参考   Reference  : IEC 61131-3:2013 §6.6.3 位串 AND / OR / XOR / NOT 语义与位宽约定
  平台   Platform   : 纯 IEC 61131-3（AND / OR / XOR / NOT / 类型转换），三平台通用
  依赖   Depends    : 仅 Standard.library（无库调用）
  分工声明 Split     : FC_DL_BitFieldExtract 为无符号位段提取属主；FC_DL_WordToIntSat
                      为整字宽（16 位整字）饱和属主；本件为任意窄位宽的有符号/零扩展，
                      三者边界：多位段拼接用前者，整字溢出饱和用中者，窄位宽符号还原用本件。
  归属 Ownership     : 本件无 TYPE 声明；常量表 DL_SEXT_LO 为本文件私有常量。
  典型用途 Use      : Modbus 双字有符号量拼装（先拼 32 位再按 16 位符号还原）、
                      12 / 16 位 ADC 原始码还原、位域字段解包。
  ------------------------------------------------------------------
  边界 Boundary     :
                      一 nWidth 越域（< 1 或 > 32）判故障并早退返回 FALSE，禁静默钳位：
                         位宽错意味着调用方拼装逻辑已错，钳位后继续会掩盖协议错位；
                      二 全部掩码由单一预计算常量表 DL_SEXT_LO 派生：
                         低位掩码 = LO[n]；高位掩码 = LO[n] XOR 全 1；符号位 = LO[n] AND NOT LO[n-1]；
                         由此消灭运行时 SHL(x, nWidth)，nWidth = 32 时不触发未定义行为；
                      三 符号扩展只在符号位为 1 时 OR 高位掩码，否则零扩展路径不受污染；
                      四 纯函数：无记忆量、无定时器、无边沿实例，每调用重算。
  错误码 Codes      :
    16#0001_064D【故障级】位宽越域（nWidth < 1 或 > 32），diOut = 0，返回 FALSE
  验收 Acceptance   :
    算法已证（脚本）：未跑 ｜ 编译器已证（三平台）：未跑
    V1 nWidth=1、bSigned=TRUE、diIn=1 → -1；diIn=0 → 0
    V2 nWidth=8、bSigned=TRUE：16#0000_00FF → -1；16#0000_007F → 127
    V3 nWidth=16、bSigned=TRUE：16#0000_8000 → -32768
    V4 nWidth=32：任意值原样返回（两种 bSigned 一致）
    V5 nWidth=0 → 0 + 码 064D + 返回 FALSE；V6 nWidth=33 → 同一处置
    V7 nWidth=4、bSigned=FALSE、diIn=16#F → 15（掩码后不扩符号）
  修订记录 Revision  :
    2026-11-21  v1.0.0  R62 首版（批 2 · 序号 4）
  ==================================================================
*)
FUNCTION FC_DL_SignExtendEx : BOOL
VAR_INPUT
    diIn    : DINT; // 待扩展值 [−]，完整 DINT 域 / the value to extend over the full DINT domain
    nWidth  : DINT; // 有效位宽 [位]，合法域 1..32 / the significant width in bits, legal one to thirty two
    bSigned : BOOL; // TRUE = 符号扩展，FALSE = 零扩展 [-] / true selects the sign extension, false the zero extension
END_VAR
VAR_OUTPUT
    diOut   : DINT;  // 扩展结果 [−] / the extended result
    eErr    : UDINT; // 错误码，0 = 正常 / the error code, zero is ok
    bError  : BOOL;  // 故障标志，故障级码同拍置位（R45 配对）/ the fault flag, raised with a fault level code
END_VAR
VAR
    udwIn   : DWORD := 16#0000_0000; // 输入位型 [位] / the input bit pattern in bits
    udwLo   : DWORD := 16#0000_0000; // 低 nWidth 位掩码 [位] / the low width mask in bits
    udwHi   : DWORD := 16#0000_0000; // 高位全 1 掩码 [位] / the high side all ones mask in bits
    udwSign : DWORD := 16#0000_0000; // 符号位单点掩码 [位] / the single bit sign mask in bits
    udwOut  : DWORD := 16#0000_0000; // 扩展后位型 [位] / the extended bit pattern in bits
END_VAR  // R64 结构补齐：VAR 段缺失的 END_VAR（门禁机械修复）
VAR CONSTANT
    DL_SEXT_MINW : DINT := 1;            // 位宽下界 [位] / the width floor in bits
    DL_SEXT_MAXW : DINT := 32;           // 位宽上界（DINT 容器位宽）[位] / the width ceiling, the DINT container width
    DL_SEXT_ALL  : DWORD := 16#FFFF_FFFF; // 全 1 常量，用于取补 [位] / the all ones constant used for the complement
    DL_SEXT_LO : ARRAY[0..32] OF DWORD := // 低 n 位掩码表（第 n 项 = 低 n 位置 1），预计算禁运行时 SHL [位] / the precomputed low width mask table
    [
        16#0000_0000, // n = 0：无有效位 / n equals zero, no significant bit
        16#0000_0001, // n = 1 / one bit
        16#0000_0003, // n = 2 / two bits
        16#0000_0007, // n = 3 / three bits
        16#0000_000F, // n = 4 / four bits
        16#0000_001F, // n = 5 / five bits
        16#0000_003F, // n = 6 / six bits
        16#0000_007F, // n = 7 / seven bits
        16#0000_00FF, // n = 8：单字节 / one byte
        16#0000_01FF, // n = 9 / nine bits
        16#0000_03FF, // n = 10 / ten bits
        16#0000_07FF, // n = 11 / eleven bits
        16#0000_0FFF, // n = 12：12 位 ADC 原始码常用 / the usual twelve bit ADC raw code width
        16#0000_1FFF, // n = 13 / thirteen bits
        16#0000_3FFF, // n = 14 / fourteen bits
        16#0000_7FFF, // n = 15 / fifteen bits
        16#0000_FFFF, // n = 16：单字 / one word
        16#0001_FFFF, // n = 17 / seventeen bits
        16#0003_FFFF, // n = 18 / eighteen bits
        16#0007_FFFF, // n = 19 / nineteen bits
        16#000F_FFFF, // n = 20 / twenty bits
        16#001F_FFFF, // n = 21 / twenty one bits
        16#003F_FFFF, // n = 22 / twenty two bits
        16#007F_FFFF, // n = 23 / twenty three bits
        16#00FF_FFFF, // n = 24 / twenty four bits
        16#01FF_FFFF, // n = 25 / twenty five bits
        16#03FF_FFFF, // n = 26 / twenty six bits
        16#07FF_FFFF, // n = 27 / twenty seven bits
        16#0FFF_FFFF, // n = 28 / twenty eight bits
        16#1FFF_FFFF, // n = 29 / twenty nine bits
        16#3FFF_FFFF, // n = 30 / thirty bits
        16#7FFF_FFFF, // n = 31 / thirty one bits
        16#FFFF_FFFF  // n = 32：整容器 / the whole container
    ];
END_VAR

// 段 1｜返回值与全部出口预置安全值（R45 四段式第一段）/ segment 1, preset every outlet to its safe value
FC_DL_SignExtendEx := FALSE; // 返回值预置假 / preset the return false
diOut := 0; // 结果预置零 [−] / preset the result zero
eErr := 16#0000_0000; // 错误码预置正常 / preset the code to ok
bError := FALSE; // 故障标志预置假 / preset the fault flag false
udwIn := 16#0000_0000; // 输入位型清零 [位] / clear the input bit pattern
udwLo := 16#0000_0000; // 低位掩码清零 [位] / clear the low mask
udwHi := 16#0000_0000; // 高位掩码清零 [位] / clear the high mask
udwSign := 16#0000_0000; // 符号掩码清零 [位] / clear the sign mask
udwOut := 16#0000_0000; // 输出位型清零 [位] / clear the output bit pattern

// 段 2｜位宽域闸：越域判故障早退（边界一，禁静默钳位）/ segment 2, the width domain gate, no silent clamping
IF (nWidth < DL_SEXT_MINW) OR (nWidth > DL_SEXT_MAXW) THEN // 位宽越域 / the width is out of the domain
    eErr := 16#0001_064D; // 故障级：位宽越域 / fault grade, the width is out of the domain
    bError := TRUE; // 同拍置故障标志（R45 配对）/ raise the fault flag on the same scan
    diOut := 0; // 确定缺省值零 [−] / the deterministic default of zero
    RETURN; // 早退，禁钳后继续（钳位会掩盖调用方的协议错位）/ early return, clamping would hide a protocol misalignment
END_IF

// 段 3｜三张掩码由单一常量表派生（边界二，无运行时移位）/ segment 3, derive all three masks from the single precomputed table
udwIn := DINT_TO_DWORD(diIn); // 输入位型接管 [位] / take the input bit pattern
udwLo := DL_SEXT_LO[nWidth]; // 低 nWidth 位掩码 [位] / the low width mask
udwHi := udwLo XOR DL_SEXT_ALL; // 高位全 1 掩码 = 低掩码取补 [位] / the high mask is the complement of the low mask
udwSign := udwLo AND (NOT DL_SEXT_LO[nWidth - DL_SEXT_MINW]); // 符号位 = 第 nWidth 位（低 n 掩码与低 n-1 掩码之差）[位] / the sign bit is the n-th bit

// 段 4｜零扩展基线：先取低 nWidth 位（两条路径共用的第一段）/ segment 4, the zero extension baseline shared by both paths
udwOut := udwIn AND udwLo; // 低 nWidth 位保留，其余清零 [位] / keep the low width bits and clear the rest

// 段 5｜符号扩展：符号位为 1 才补高位全 1（边界三）/ segment 5, the sign extension only when the sign bit is set
IF bSigned THEN // 调用方要求符号扩展 / the caller asked for the sign extension
    IF (udwOut AND udwSign) <> 16#0000_0000 THEN // 符号位为 1 / the sign bit is set
        udwOut := udwOut OR udwHi; // 高位补全 1（nWidth = 32 时 udwHi 为零，等价原样返回）/ fill the high side, the width of thirty two yields a zero high mask and passes the value through
    END_IF
END_IF

// 段 6｜统一出口（位型还原为有符号结果）/ segment 6, the unified outlet
diOut := DWORD_TO_DINT(udwOut); // 位型还原 [−] / reinterpret the bit pattern as a signed value
FC_DL_SignExtendEx := TRUE; // 返回成功 / return success
END_FUNCTION

(* ---- FC_DL_SortIndexInt.st ---- *)
// ==============================================================================
// 组件名 Component  : FC_DL_SortIndexInt
// 分类   Category   : DL_Base
// 前缀   Naming     : FC_DL_ ｜ b/n/f 类型前缀制（R265）
// 版本   Version    : 1.0.0
// 复杂度 Complexity  : 中
// 功能   Purpose    : INT 数组稳定索引排序：输出按值排序后的原下标排列，
//                      不改 arrSrc（只读纪律）；bDesc = FALSE 升序 /
//                      TRUE 降序；等值元素保持原下标先后（稳定性判据 =
//                      严格比较 + 不交换等值对）。nUsed 钳位 [0, 64]。
// 开源溯源 Origin    : 道莅原创（与 DL_MathData 的 FC_DL_SortIndexLReal
//                      同族自研语义，索引间接排序实现，零代码复制）
// 许可证 License    : MIT
// 参考   Reference  : IEC 61131-3:2013 §6.6.4 FOR / WHILE 遍历语义
// 平台   Platform   : 纯 IEC 61131-3（FOR / WHILE / 比较 / 数组），三平台通用
// 依赖   Depends    : 无（零委托、零库件）
// 分工声明 Split     : FC_DL_SortIndexLReal（LREAL 版索引排序）为本件同族
//                      件，两件类型口径不同、语义同源，互引声明（R216）；
//                      本件只出索引排列不改数据，读写纪律与彼件一致。
// 归属 Ownership     : 本件无 TYPE 声明；全部引脚为 IEC 标准原生类型。
// ------------------------------------------------------------------
// 边界 Boundary     :
//   一 计数域闸：nUsed < 0 → 恒等索引早退合法返回（nSorted = 0）；nUsed
//      > 64 → 钳 64 续排（信息级语义，本件无 eErr 出口，钳位场景出口与
//      正常截断排序同形、无独立通道可承载，不另设码，R90 反证句）；
//   二 稳定性判据写死下标序：升序用严格大于、降序用严格小于前移，相等
//      元素不交换（插入序即下标序），升 / 降两向稳定性自证；
//   三 索引写出前已证在 [0, nUse-1] 内（arrIdx 恒等预置 + 插入原地移动），
//      回钳量不复判越界（R241）；
//   四 WHILE 护栏计数 nGuard（上界 32000，远大于最坏比较次数 64*63/2 =
//      2016，且 nGuard 为 INT 不溢出），护栏命中强制退出内层（结构性
//      不可达兜底，不静默死循环）；
//   五 INT 元素无非有限面（NaN / Inf 不适用于整型），非有限闸 N/A；
//   六 nUsed = 0 / 1 退化直返恒等索引（arrIdx[i] = i），bValid = TRUE；
//   七 纯函数：无记忆量、无定时器、无边沿实例，每调用重算；
//   八 无除法；无全局、无外部变量、无物理地址。
// 错误码 Codes      :
//   16#0001_0746【信息级】nUsed 越域已钳位（< 0 恒等早退，> 64 钳 64 续排）
//   注：本件引脚契约按任务定稿无独立 eErr 出口，钳位语义为文档级。
// 验收 Acceptance   :
//   算法已证（脚本）：未跑 ｜ 编译器已证（三平台）：未跑
//   V1 值 3/1/2 → 升序索引 1/2/0；V2 值 2/2/1 → 升序索引 2/0/1（稳定性）
//   V3 值 2/2/1 → 降序索引 0/1/2（降序稳定性同向自证）
//   V4 nUsed = 0 / 1 → 恒等索引；V5 nUsed = 100 → 钳 64 续排
//   V6 调用后 arrSrc 原样（只读纪律）
// 修订记录 Revision  :
//   2026-11-22  v1.0.0  R65 首版（批 2 · 序号 5）
// ==============================================================================
FUNCTION FC_DL_SortIndexInt : BOOL
VAR_IN_OUT
    arrSrc : ARRAY[0..63] OF INT; // 待排序数值 [-]，只读纪律（不改调用方数组）/ the values to sort, read only
END_VAR
VAR_INPUT
    nUsed : INT := 0;            // 参与排序个数 [个]，合法域 0..64 / the count, legal zero to sixty four
    bDesc : BOOL := FALSE;       // 降序开关 [-]，FALSE 升序 / the descending switch, false is ascending
END_VAR
VAR_OUTPUT
    arrIdx  : ARRAY[0..63] OF INT; // 排序后索引排列（arrIdx[0] 为极值原下标）/ the sorted index permutation
    nSorted : INT;               // 实际排序个数 [个] / the actually sorted count
    bValid  : BOOL;              // 结果可用 [-] / the result usable flag
END_VAR
VAR
    k       : INT;               // 外层插入索引 [下标] / the outer insertion index
    m       : INT;               // 内层前移索引 [下标] / the inner shifting index
    nUse    : INT;               // 钳位后的个数 [个] / the clamped count
    nKey    : INT;               // 待插元素原下标暂存 [下标] / the key original index in staging
    nKeyVal : INT;               // 待插元素值暂存 [-] / the key value in staging
    nGuard  : INT;               // 护栏计数 [次] / the guard counter
END_VAR
VAR CONSTANT
    DL_SII_NMAX : INT := 64;     // 排序容量上界 [个]，与数组容量一致 / the capacity aligned with the array
    DL_SII_GMAX : INT := 32000;  // 护栏计数上界 [次]，大于最坏比较次数 2016 且 INT 不溢出 / the guard bound above the worst case
END_VAR

// 段 1｜返回值与全部出口预置 + 索引数组恒等预置（R45 / R254）/ segment 1, the preset and the identity preset
FC_DL_SortIndexInt := FALSE;     // 返回值预置假 / preset the return false
nSorted := 0;                    // 排序个数预置零 [个] / preset the sorted count zero
bValid  := FALSE;                // 有效标志预置假 / preset the validity false
nUse    := 0;                    // 个数预置零 [个] / preset the count zero
nKey    := 0;                    // 键下标预置零 [下标] / preset the key index zero
nKeyVal := 0;                    // 键值预置零 / preset the key value zero
nGuard  := 0;                    // 护栏预置零 [次] / preset the guard zero
FOR k := 0 TO DL_SII_NMAX - 1 DO // 索引数组全量预置恒等 / preset the index array to the identity
    arrIdx[k] := k;              // 恒等索引 / the identity index
END_FOR

// 段 2｜计数域闸（边界一：负数恒等早退，超容量钳位续排）/ segment 2, the count domain gate
IF nUsed < 0 THEN                // 负数非法 / a negative count
    bValid := TRUE;              // 空排列合法（arrIdx 已全量恒等）/ an empty permutation is legal
    FC_DL_SortIndexInt := TRUE;  // 返回成功 / return success
    RETURN;                      // 早退（信息级 0746 语义，文档级）/ early return
END_IF
nUse := nUsed;                   // 域内接管 / take the count
IF nUse > DL_SII_NMAX THEN       // 超容量 / above the capacity
    nUse := DL_SII_NMAX;         // 钳到容量（信息级 0746 语义）/ clamp to the capacity
END_IF

// 段 3｜稳定插入排序（索引间接，严格比较保稳定，边界二；护栏防死循环，边界四）/ segment 3, the stable insertion sort on the indices
FOR k := 1 TO nUse - 1 DO        // 有界外层 / the bounded outer loop
    nKey := arrIdx[k];           // 待插元素原下标 / the key original index
    nKeyVal := arrSrc[nKey];     // 待插元素值 / the key value
    m := k - 1;                  // 内层从前一位置起 / the inner scan starts here
    nGuard := 0;                 // 护栏清零 / reset the guard
    WHILE (m >= 0) AND (((NOT bDesc) AND (arrSrc[arrIdx[m]] > nKeyVal)) OR (bDesc AND (arrSrc[arrIdx[m]] < nKeyVal))) DO // 前驱按序更极才前移（严格比较，等值不交换，稳定性自证）/ shift while the predecessor is strictly more extreme
        arrIdx[m + 1] := arrIdx[m]; // 索引后移一位 / shift the index right
        m := m - 1;              // 内层前移 / step the inner scan left
        nGuard := nGuard + 1;    // 护栏计数推进 / advance the guard
        IF nGuard > DL_SII_GMAX THEN // 护栏命中（结构性不可达兜底）/ the guard tripped
            m := -1;             // 强制退出内层（不置码，结构兜底）/ force the inner loop out
        END_IF
    END_WHILE
    arrIdx[m + 1] := nKey;       // 键落位（m+1 已证在 [0, k] 内，边界三）/ the key lands with a proven bound
END_FOR

// 段 4｜出口（nUse = 0/1 时 arrIdx 已为恒等，边界六）/ segment 4, the outlet with the degenerate identity
nSorted := nUse;                 // 排序个数出口 [个] / the sorted count outlet
bValid := TRUE;                  // 结果可用 / the result usable
FC_DL_SortIndexInt := TRUE;      // 返回成功 / return success
END_FUNCTION
